(* IEC 61131-3 sources: FibonacciChallenge/Class/SafetyManager (part 3) *)

        pPDOElement^.PDO_ID                 := PDO_ID;
        pPDOElement^.Length                 := Length;
        pPDOElement^.ThisDomainsRole        := SourceDest_IsDest;

        pPDOElement^.SourceInfo.SafetyNbr   := 0;
        pPDOElement^.SourceInfo.DomainNr    := SourceDomain;
        pPDOElement^.SourceInfo.PathLen     := SourcePathLen;
        pPDOElement^.SourceInfo.pPath$pVoid := To_StdLib.Malloc(size:= SourcePathLen);
        if pPDOElement^.SourceInfo.pPath then
          _memcpy(ptr1:=pPDOElement^.SourceInfo.pPath, ptr2:=pSourcePath, cntr:=SourcePathLen);
        else
          LogError("@0464 (SafetyManager::IsAffectedByPDO) Failed to allocate memory for PDO path info");
          ClassState := -1;
          return;
        end_if;

        pPDOElement^.DestInfo.SafetyNbr     := pSafetyNbr^;
        pPDOElement^.DestInfo.DomainNr      := DestDomain;
        pPDOElement^.DestInfo.PathLen       := DestPathLen;
        pPDOElement^.DestInfo.pPath$pVoid   := To_StdLib.Malloc(size:= DestPathLen);
        if pPDOElement^.DestInfo.pPath then
          _memcpy(ptr1:=pPDOElement^.DestInfo.pPath, ptr2:=pDestPath, cntr:=DestPathLen);
        else
          LogError("@0464 (SafetyManager::IsAffectedByPDO) Failed to allocate memory for PDO path info");
          ClassState := -1;
          return;
        end_if;

        pPDOElement^.pSafety              := pDestSafety;

        // if we're the master, we may also route interfaceframes
        if IsInterfaceFrame then

          // search for the source of this PDO
          pHelpManaging := pFirstManagingInterfaceComponent;
          while pHelpManaging do
            if (To_StdLib.MemCmp(pHelpManaging^.pModulePath, pSourcePath, SourcePathLen) = 0) then
              exit;
            else
              pHelpManaging := pHelpManaging^.pNext;
            end_if;
          end_while;

          pPDOElement^.pManagingSource := pHelpManaging;
        end_if;

        if pPDOElement^.pManagingSource then

          // if the module is marked as optional and the PDO is not optional => the module is also not optional
          if pPDOElement^.pManagingSource^.InfoBits.IsOptional & (PDOInfo.IsOptional = FALSE) then
            pPDOElement^.pManagingSource^.InfoBits.IsOptional  := FALSE;
          end_if;

          // check if we can recycle the memory of another DO (if this data is already transferred to this managing module
          pRecyclePDO := CheckPDORecycle(SourceDest_IsSource, pPDOElement);

          // only if there is enough space or we already have a memory
          if pRecyclePDO | ((pPDOElement^.pManagingSource^.PDOReadMemUsed + pPDOElement^.Length) <= pPDOElement^.pManagingSource^.PDOReadMemAvailable) then
            if IsInterfaceFrame then
              pPDOElement^.SourceInfo.SafetyNbr   := (GetIFInfoByCRC(InterfaceCRC, #TempOffset, #TempLen))$HDINT;
              if TempLen = Length then
                // get the place in the memory of the source managing module
                pPDOElement^.SourceInfo.pPDOMem       := pPDOElement^.pManagingSource^.pPDOReadSpace + TempOffset;
                pPDOElement^.SourceInfo.pPDOMemDPRAM  := pPDOElement^.pManagingSource^.pPDOReadSpaceDPRAM + TempOffset;

                pPDOElement^.SourceInfo.HandlePDODPRAM := pPDOElement^.pManagingSource^.ud_HandlePDOReadSpaceDPRAM;
                pPDOElement^.SourceInfo.OffsetPDODPRAM := TempOffset;

                // if we need new memory, tell the managing module
                if (TempOffset + Length) > pPDOElement^.pManagingSource^.PDOReadMemUsed then
                  pPDOElement^.pManagingSource^.PDOReadMemUsed := TempOffset + Length;

                  MyPara.uiCmd := CMD_SM_PDO_MEM_USAGE_RD;
                  MyPara.aPara[0] := pPDOElement^.pManagingSource^.PDOReadMemUsed$DINT;
                  pPDOElement^.pManagingSource^.pThis^.NewInst(#MyPara, #MyResult);
                end_if;

                MyPara.uiCmd := CMD_SM_ADD_INPUT_PDO;
                MyPara.aPara[0] := pPDOElement^.SourceInfo.pPDOMem$DINT;
                MyPara.aPara[1] := pPDOElement^.SourceInfo.pPDOMemDPRAM$DINT;
                MyPara.aPara[2] := pPDOElement^.SourceInfo.SafetyNbr$DINT;
                MyPara.aPara[3] := Length;
                MyPara.aPara[4] := PDOInfo.IsOptional;
                MyPara.aPara[5] := pPDOElement^.SourceInfo.HandlePDODPRAM$DINT; // Needed for Payload Support
                MyPara.aPara[6] := pPDOElement^.SourceInfo.OffsetPDODPRAM$DINT; // Needed for Payload Support
                MyPara.aPara[7] := 0;// target offset (not necessary here)
                MyPara.aPara[8] := SM_IF_VALIDITY_MARK$DINT;
                MyPara.aPara[9] := TRUE;

                pDestSafety^.pThis^.NewInst(#MyPara, #MyResult);
              else
                LogError("@0469 (SafetyManager::IsAffectedByPDO) Length of interface frames doesn't match the local configuration");
              end_if;

            else
              if pRecyclePDO then
                pPDOElement^.SourceInfo.pPDOMem       := pRecyclePDO^.SourceInfo.pPDOMem;
                pPDOElement^.SourceInfo.pPDOMemDPRAM  := pRecyclePDO^.SourceInfo.pPDOMemDPRAM;
              else
                pPDOElement^.SourceInfo.pPDOMem       := pPDOElement^.pManagingSource^.pPDOReadSpace + pPDOElement^.pManagingSource^.PDOReadMemUsed;
                pPDOElement^.SourceInfo.pPDOMemDPRAM  := pPDOElement^.pManagingSource^.pPDOReadSpaceDPRAM + pPDOElement^.pManagingSource^.PDOReadMemUsed;

                // if we need new memory, tell the managing module
                pPDOElement^.pManagingSource^.PDOReadMemUsed += pPDOElement^.Length;

                MyPara.uiCmd := CMD_SM_PDO_MEM_USAGE_RD;
                MyPara.aPara[0] := pPDOElement^.pManagingSource^.PDOReadMemUsed$DINT;
                pPDOElement^.pManagingSource^.pThis^.NewInst(#MyPara, #MyResult);
              end_if;
            end_if;
          else
            // we add the memory anyway to show the user how much he would need
            pPDOElement^.pManagingSource^.PDOReadMemUsed += pPDOElement^.Length;

            MyPara.uiCmd := CMD_SM_PDO_MEM_USAGE_RD;
            MyPara.aPara[0] := pPDOElement^.pManagingSource^.PDOReadMemUsed$DINT;
            pPDOElement^.pManagingSource^.pThis^.NewInst(#MyPara, #MyResult);

            LogError("@046B (SafetyManager::IsAffectedByPDO) Not enough read memory to map all PDOs");
            return;
          end_if;
        else

          LogError("@046C (SafetyManager::IsAffectedByPDO) Couldn't find source managing module for PDO");
          return;
        end_if;

        PDOElementNo += 1;
      else
        pSourceDest^ := SourceDest_IsForwarder;

        // if source and destination are not in this domain, is it a bifurcation or a linear forwarding?
        pPDOElement^.PDO_ID                 := PDO_ID;
        pPDOElement^.Length                 := Length;
        pPDOElement^.ThisDomainsRole        := SourceDest_IsForwarder;

        pPDOElement^.SourceInfo.DomainNr    := SourceDomain;
        pPDOElement^.SourceInfo.PathLen     := SourcePathLen;
        pPDOElement^.SourceInfo.pPath$pVoid := To_StdLib.Malloc(size:= SourcePathLen);
        if pPDOElement^.SourceInfo.pPath then
          _memcpy(ptr1:=pPDOElement^.SourceInfo.pPath, ptr2:=pSourcePath, cntr:=SourcePathLen);
        else
          LogError("@0464 (SafetyManager::IsAffectedByPDO) Failed to allocate memory for PDO path info");
          ClassState := -1;
          return;
        end_if;

        pPDOElement^.DestInfo.DomainNr      := DestDomain;
        pPDOElement^.DestInfo.PathLen       := DestPathLen;
        pPDOElement^.DestInfo.pPath$pVoid   := To_StdLib.Malloc(size:= DestPathLen);
        if pPDOElement^.DestInfo.pPath then
          _memcpy(ptr1:=pPDOElement^.DestInfo.pPath, ptr2:=pDestPath, cntr:=DestPathLen);
        else
          LogError("@0464 (SafetyManager::IsAffectedByPDO) Failed to allocate memory for PDO path info");
          ClassState := -1;
          return;
        end_if;

        // initialize with invalid;
        CopyCmdIndex := -1;

        // if we're the master, we may also route interfaceframes
        if IsInterfaceFrame then

          // search for the source of this PDO
          pHelpManaging := pFirstManagingInterfaceComponent;
          while pHelpManaging do
            if (To_StdLib.MemCmp(pHelpManaging^.pModulePath, pSourcePath, SourcePathLen) = 0) then
              exit;
            else
              pHelpManaging := pHelpManaging^.pNext;
            end_if;
          end_while;

          pPDOElement^.pManagingSource := pHelpManaging;
        end_if;

        if pPDOElement^.pManagingSource then

          // if the module is marked as optional and the PDO is not optional => the module is also not optional
          if pPDOElement^.pManagingSource^.InfoBits.IsOptional & (PDOInfo.IsOptional = FALSE) then
            pPDOElement^.pManagingSource^.InfoBits.IsOptional  := FALSE;
          end_if;

          // check if we can recycle the memory of another DO (if this data is already transferred to this managing module
          pRecyclePDO := CheckPDORecycle(SourceDest_IsSource, pPDOElement);

          if pRecyclePDO | ((pPDOElement^.pManagingSource^.PDOReadMemUsed + pPDOElement^.Length) <= pPDOElement^.pManagingSource^.PDOReadMemAvailable) then
            if pRecyclePDO then
              pPDOElement^.SourceInfo.pPDOMem       := pRecyclePDO^.SourceInfo.pPDOMem;
              pPDOElement^.SourceInfo.pPDOMemDPRAM  := pRecyclePDO^.SourceInfo.pPDOMemDPRAM;
            else
              pPDOElement^.SourceInfo.pPDOMem       := pPDOElement^.pManagingSource^.pPDOReadSpace + pPDOElement^.pManagingSource^.PDOReadMemUsed;
              pPDOElement^.SourceInfo.pPDOMemDPRAM  := pPDOElement^.pManagingSource^.pPDOReadSpaceDPRAM + pPDOElement^.pManagingSource^.PDOReadMemUsed;
              pPDOElement^.pManagingSource^.PDOReadMemUsed += pPDOElement^.Length;

              MyPara.uiCmd := CMD_SM_PDO_MEM_USAGE_RD;
              MyPara.aPara[0] := pPDOElement^.pManagingSource^.PDOReadMemUsed$DINT;
              pPDOElement^.pManagingSource^.pThis^.NewInst(#MyPara, #MyResult);
            end_if;
          else
            // we add the memory anyway to show the user how much he would need
            pPDOElement^.pManagingSource^.PDOReadMemUsed += pPDOElement^.Length;

            MyPara.uiCmd := CMD_SM_PDO_MEM_USAGE_RD;
            MyPara.aPara[0] := pPDOElement^.pManagingSource^.PDOReadMemUsed$DINT;
            pPDOElement^.pManagingSource^.pThis^.NewInst(#MyPara, #MyResult);

            LogError("@046B (SafetyManager::IsAffectedByPDO) Not enough read memory to map all PDOs");
            return;
          end_if;
        else
          LogError("@046C (SafetyManager::IsAffectedByPDO) Couldn't find source managing module for PDO");
          return;
        end_if;

        // if we're the master, we may also route interfaceframes
        if IsInterfaceFrame then
          // search for the destination of this PDO
          pHelpManaging := pFirstManagingInterfaceComponent;
          while pHelpManaging do
            if (To_StdLib.MemCmp(pHelpManaging^.pModulePath, pDestPath, DestPathLen) = 0) then
              exit;
            else
              pHelpManaging := pHelpManaging^.pNext;
            end_if;
          end_while;

          pPDOElement^.pManagingDest := pHelpManaging;
        end_if;

        if pPDOElement^.pManagingDest then

          // if the module is marked as optional and the PDO is not optional => the module is also not optional
          if pPDOElement^.pManagingDest^.InfoBits.IsOptional & (PDOInfo.IsOptional = FALSE) then
            pPDOElement^.pManagingDest^.InfoBits.IsOptional  := FALSE;
          end_if;

          if pPDOElement^.pManagingDest = pPDOElement^.pManagingSource then
            LogError("@0470 (SafetyManager::IsAffectedByPDO) In PDO Forwarding a domain can't be the source and the destination!");
          end_if;

          // check if we can recycle the memory of another DO (if this data is already transferred to this managing module
          pRecyclePDO := CheckPDORecycle(SourceDest_IsDest, pPDOElement);

          if pRecyclePDO | ((pPDOElement^.pManagingDest^.PDOWriteMemUsed + pPDOElement^.Length) <= pPDOElement^.pManagingDest^.PDOWriteMemAvailable) then

            // if we can't use the copy command
            if b_SafetyOnLocalCDIAS then
              // remember the pointer to the memory to copy it manually in rt postscan method
              if pRecyclePDO then
                // this PDO is already in the memory of the managing node, we don't have to copy it again
                pPDOElement^.DestInfo.pPDOMem := NIL;//pRecyclePDO^.SourceInfo.pPDOMem;
              else
                pPDOElement^.DestInfo.pPDOMem := pPDOElement^.pManagingDest^.pPDOWriteSpace + pPDOElement^.pManagingDest^.PDOWriteMemUsed;
              end_if;
            else
              if pRecyclePDO then
                // this PDO is already in the memory of the managing node, we don't have to copy it again
                pPDOElement^.DestInfo.pPDOMemDPRAM := NIL;//pRecyclePDO^.DestInfo.pPDOMemDPRAM;
              else
                pPDOElement^.DestInfo.pPDOMemDPRAM := pPDOElement^.pManagingDest^.pPDOWriteSpaceDPRAM + pPDOElement^.pManagingDest^.PDOWriteMemUsed;
              end_if;

              CopyCmdIndex := GetNewMovDO();
              if CopyCmdIndex < 0 then
                pPDOElement^.DestInfo.pPDOMem := pPDOElement^.pManagingDest^.pPDOWriteSpace + pPDOElement^.pManagingDest^.PDOWriteMemUsed;
                LogError("@0465 (SafetyManager::IsAffectedByPDO) Failed to install copy command => PDO is beeing copied in RT");
              else
                aCopyCmds[CopyCmdIndex].pSettings^.ud_AddressDest := pPDOElement^.DestInfo.pPDOMemDPRAM$UDINT;
                aCopyCmds[CopyCmdIndex].pSettings^.ui_ByteCnt     := pPDOElement^.Length;
              end_if;
            end_if;

            // if we need new memory, tell the managing module
            if pRecyclePDO = NIL then
              pPDOElement^.pManagingDest^.PDOWriteMemUsed += pPDOElement^.Length;

              MyPara.uiCmd := CMD_SM_PDO_MEM_USAGE_WR;
              MyPara.aPara[0] := pPDOElement^.pManagingDest^.PDOWriteMemUsed$DINT;
              pPDOElement^.pManagingDest^.pThis^.NewInst(#MyPara, #MyResult);
            end_if;
          else
            // we add the memory anyway to show the user how much he would need
            pPDOElement^.pManagingDest^.PDOWriteMemUsed += pPDOElement^.Length;

            MyPara.uiCmd := CMD_SM_PDO_MEM_USAGE_WR;
            MyPara.aPara[0] := pPDOElement^.pManagingDest^.PDOWriteMemUsed$DINT;
            pPDOElement^.pManagingDest^.pThis^.NewInst(#MyPara, #MyResult);

            LogError("@0466 (SafetyManager::IsAffectedByPDO) Not enough write memory to map all PDOs");
            return;
          end_if;
        else
          LogError("@0467 (SafetyManager::IsAffectedByPDO) Couldn't find destination managing module for PDO");
          return;
        end_if;

        pPDOElement^.CopyCmdIndex := CopyCmdIndex;

        PDOElementNo += 1;
      end_if;

    end_if;
  end_if;

END_FUNCTION

FUNCTION SafetyManager::GetDestManagingOfDO
  VAR_INPUT
    pDO 	: ^SafetyCDIAS_Base::SDOHeader;
  END_VAR
  VAR_OUTPUT
    pDestManaging 	: ^t_ManagingComponent;
  END_VAR
  VAR
    pHelpManaging 	          : ^t_ManagingComponent;
    pAddDynSlaveRsp           : ^t_AddDynSlaveRsp;
    pRemDynSlaveRsp           : ^t_RemDynSlaveRsp;
    pHelpConfig               : ^t_CfgListElem;
    pHelpConnection           : ^t_FSoEConnectionDetails;
    MyPara                    : CmdStruct;
    MyResult                  : results;
    i                         : USINT;
    b_ConnectionAlreadyExists : BOOL;
  END_VAR

  pDestManaging := NIL;

  // maybe it's one of the interface domains
  pHelpManaging := pFirstManagingInterfaceComponent;
  while pHelpManaging do
    if (pHelpManaging^.FlexCon.SafetyNumber = pDO^.DstAdr) then
      if (pDO^.StdHeader.Typ.Response) & ((pDO^.StdHeader.Cmd = SM_SDO_COMMAND_ADD_DYN_SLAVE) | (pDO^.StdHeader.Cmd = SM_SDO_COMMAND_REMOVE_DYN_SLAVE)) then

        // if the initialisation of the class is not finished or failed
        if (sFlexCon.Role <> _NoFlexCon) & (ClassState <> 1) then
          // don't forward add or remove dyn slave requests. otherwise the order in the managing module is likely to be wrong if flexcon is used in combination with interface frames.
          return;
        end_if;

        if (pDO^.StdHeader.Cmd = SM_SDO_COMMAND_ADD_DYN_SLAVE) then
          pAddDynSlaveRsp := pDO$^t_AddDynSlaveRsp;

          // if it was successful and we have a safety host module pointer => try to install the PDO
          if (pAddDynSlaveRsp^.Retcode = 0) & sFlexCon.pSafetyHost then
#ifdef SAFETY_DEBUG_LOGGING_ACTIVATED
            LogError("@DBG AddDynSlave Response detected in SafetyManager of Host (succeeded)");
#endif

            // install the access to the next free memory on the VBC

            // we're the host => search for the FSoE connection with the host flags
            pHelpConfig := pConfigs;
            while pHelpConfig do
              pHelpConnection := pHelpConfig^.pFirstFSoEConnection;
              while pHelpConnection do
                if ((pHelpConnection^.Flags AND SM_FLAGS_FLEXCON_MASK) = SM_FLAGS_FLEXCON_HOST) &   // check if it's the right kind of connection
//                   (pHelpConnection^.InternalConnectionState =  FCS_RESET)               &          // check if it's still free
                   (pHelpConnection^.MasterReadOffset  = pAddDynSlaveRsp^.SafeOutOffset) &          // check if offsets and lengths match
                   (pHelpConnection^.MasterWriteOffset = pAddDynSlaveRsp^.SafeInOffset)  &
                   (pHelpConnection^.MasterReadSize    = pAddDynSlaveRsp^.SafeOutLength) &
                   (pHelpConnection^.MasterWriteSize   = pAddDynSlaveRsp^.SafeInLength) then

#ifdef SAFETY_DEBUG_LOGGING_ACTIVATED
                  LogValue(pString:="@DBG HOST: Found FSoE Connection of FlexConHost to install the cyclic PDO Routing between 0x{0} local and 0x{1} at Node", Value:=pHelpConnection^.OwnerSafetyNbr, Value2:=pHelpManaging^.FlexCon.SafetyNumber);
#endif

                  // remember if we already had this connection before
                  b_ConnectionAlreadyExists := pHelpManaging^.FlexCon.pCopyCmd <> NIL;

                  if b_ConnectionAlreadyExists = FALSE then
                    pHelpManaging^.FlexCon.WriteOffset:= pHelpManaging^.PDOWriteMemUsed$UINT;
                    pHelpManaging^.FlexCon.WriteLen   := pHelpConnection^.MasterReadSize;
                  end_if;

                  // GET THE DATA FROM THE SCP TO THE VBC

                  MyPara.uiCmd := CMD_SM_ADD_OUTPUT_PDO;
//                      MyPara.aPara[0] := 1;  not used // mark as interface frame PDO
                  sFlexCon.pSafetyHost^.pThis^.NewInst(#MyPara, #MyResult);

  //                  pPDOElement^.SourceInfo.pPDOMem       := MyResult.aData[0]$^USINT;
  //                  pPDOElement^.SourceInfo.pPDOMemDPRAM  := MyResult.aData[4]$^USINT;
  //                  pPDOElement^.SourceInfo.HandlePDODPRAM:= MyResult.aData[8]$UDINT;   // Needed for Payload Support
  //                  pPDOElement^.SourceInfo.OffsetPDODPRAM:= MyResult.aData[12]$UDINT;  // Needed for Payload Support

                  // check if we already have a copy pointer
                  if pHelpManaging^.FlexCon.pCopyCmd then
                    pHelpManaging^.FlexCon.pCopyCmd^.pSource  := MyResult.aData[0]$^USINT + pHelpConnection^.MasterReadOffset;
                    pHelpManaging^.FlexCon.pCopyCmd^.pDest    := pHelpManaging^.pPDOWriteSpace + pHelpManaging^.FlexCon.WriteOffset;
                    pHelpManaging^.FlexCon.pCopyCmd^.Size     := pHelpManaging^.FlexCon.WriteLen;
                  else
                    // create a new
                    if FSoECopyCmdNo < MAX_FSOE_CONNECTIONS then
                      aFSoECopyCmds[FSoECopyCmdNo].pSource  := MyResult.aData[0]$^USINT + pHelpConnection^.MasterReadOffset;
                      aFSoECopyCmds[FSoECopyCmdNo].pDest    := pHelpManaging^.pPDOWriteSpace + pHelpManaging^.FlexCon.WriteOffset;
                      aFSoECopyCmds[FSoECopyCmdNo].Size     := pHelpManaging^.FlexCon.WriteLen;
                      pHelpManaging^.FlexCon.pCopyCmd := #aFSoECopyCmds[FSoECopyCmdNo];
                      FSoECopyCmdNo                         += 1;
                    else
                      LogValue("@0493 (SafetyManager::GetDestManagingOfDO) Maximum limit of allowed FSoE connections exceeded (0x{0})", Value:=MAX_FSOE_CONNECTIONS);
                    end_if;
                  end_if;

                  if b_ConnectionAlreadyExists = FALSE then
                    pHelpManaging^.PDOWriteMemUsed += pHelpManaging^.FlexCon.WriteLen;
                    MyPara.uiCmd    := CMD_SM_PDO_MEM_USAGE_WR;
                    MyPara.aPara[0] := pHelpManaging^.PDOWriteMemUsed$DINT;
                    pHelpManaging^.pThis^.NewInst(#MyPara, #MyResult);

                    pHelpManaging^.FlexCon.ReadOffset := pHelpManaging^.PDOReadMemUsed$UINT;
                    pHelpManaging^.FlexCon.ReadLen    := pHelpConnection^.MasterWriteSize;
                  end_if;

                  // HOW TO GET DATA FROM THE VBC TO THE SCP

                  MyPara.uiCmd := CMD_SM_ADD_INPUT_PDO;
                  MyPara.aPara[0] := (pHelpManaging^.pPDOReadSpace + pHelpManaging^.FlexCon.ReadOffset)$DINT;
                  MyPara.aPara[1] := 0;
                  MyPara.aPara[2] := pHelpManaging^.FlexCon.SafetyNumber$DINT;
                  MyPara.aPara[3] := pHelpManaging^.FlexCon.ReadLen;
                  MyPara.aPara[4] := 0;
                  MyPara.aPara[5] := 0;
                  MyPara.aPara[6] := 0;
                  MyPara.aPara[7] := pHelpConnection^.MasterWriteOffset;
                  MyPara.aPara[8] := SM_IF_VALIDITY_MARK$DINT;
                  MyPara.aPara[9] := FALSE; // no interface frame => needed to reuse the same input PDO at the module

                  if sFlexCon.pSafetyHost^.pThis^.NewInst(#MyPara, #MyResult) = ERROR then
                    LogError(e_msg:="@05DE (SafetyManager::GetDestManagingOfDO) Failed to add FlexCon PDO to safe CPU PDO input buffer (Host side)");
                  end_if;

                  // check if we already have a input pdo pointer
                  if pHelpManaging^.FlexCon.pInputPdo then
                    pHelpManaging^.FlexCon.pInputPdo^.pSafety := sFlexCon.pSafetyHost;
                    pHelpManaging^.FlexCon.pInputPdo^.pMem    := MyPara.aPara[0];
                  else
                    if FSoEInputPDONo < MAX_FSOE_CONNECTIONS then
                      aFSoEInputPDOs[FSoEInputPDONo].pSafety    := sFlexCon.pSafetyHost;
                      aFSoEInputPDOs[FSoEInputPDONo].pMem       := MyPara.aPara[0];
                      pHelpManaging^.FlexCon.pInputPdo          := #aFSoEInputPDOs[FSoEInputPDONo];
                      FSoEInputPDONo += 1;
                    else
                      LogValue("@0490 (SafetyManager::GetDestManagingOfDO) Maximum limit of allowed FSoE input Frames exceeded (0x{0})", Value:=MAX_FSOE_CONNECTIONS);
                    end_if;
                  end_if;

#ifdef SAFETY_DEBUG_LOGGING_ACTIVATED
  #pragma message("RamAnd 20.11.2014 16:41 \ testweise mapping loggen")
                  LogValue("@DBG (SafetyManager::GetDestManagingOfDO) Mng => Modul: Wr Offset Modul: 0x{0}, Rd Offset Mng: 0x{1}, Größe: 0x{2}", Value:=pHelpConnection^.MasterWriteOffset, Value2:=pHelpManaging^.FlexCon.ReadOffset, Value3:=pHelpManaging^.FlexCon.ReadLen);
                  LogValue("@DBG (SafetyManager::GetDestManagingOfDO) Modul => Mng: Rd Offset Modul: 0x{0}, Wr Offset Mng: 0x{1}, Größe: 0x{2}", Value:=pHelpConnection^.MasterReadOffset, Value2:=pHelpManaging^.FlexCon.WriteOffset, Value3:=pHelpManaging^.FlexCon.WriteLen);
#endif

                  if b_ConnectionAlreadyExists = FALSE then
                    pHelpManaging^.PDOReadMemUsed += pHelpManaging^.FlexCon.ReadLen;

                    MyPara.uiCmd := CMD_SM_PDO_MEM_USAGE_RD;
                    MyPara.aPara[0] := pHelpManaging^.PDOReadMemUsed$DINT;
                    pHelpManaging^.pThis^.NewInst(#MyPara, #MyResult);
                  end_if;

                  // mark the connection as established
//                  pHelpConnection^.InternalConnectionState := FCS_CONNECTION;

                  // remember the connection if it's connected
                  pHelpManaging^.FlexCon.pFSoEConnection := pHelpConnection;

                  // we got our connection, stop cycling through the rest of the configurations
                  pDestManaging := pHelpManaging;
                  return;
                end_if;

                pHelpConnection := pHelpConnection^.pNext;
              end_while;
              pHelpConfig := pHelpConfig^.pNext;
            end_while;
          else
            LogValue(pString:="@05DF (SafetyManager::GetDestManagingOfDO) AddDynSlave Response detected in SafetyManager of Host (failed with retcode 0x{0})", Value:=pAddDynSlaveRsp^.Retcode);
          end_if;
        else
          pRemDynSlaveRsp := pDO$^t_RemDynSlaveRsp;

          if pRemDynSlaveRsp^.Retcode = 0 then
#ifdef SAFETY_DEBUG_LOGGING_ACTIVATED
            LogError("@DBG RemoveDynSlave Response detected in SafetyManager of Host (succeeded)");
#endif
            if pHelpManaging^.FlexCon.pFSoEConnection then
              // remove the InputPDO from the Safety CPU
              if pHelpManaging^.FlexCon.pInputPdo & pHelpManaging^.FlexCon.pInputPdo^.pMem & pHelpManaging^.FlexCon.pInputPdo^.pSafety then
                // unregister this PDO
                MyPara.uiCmd := CMD_SM_REMOVE_INPUT_PDO;
                MyPara.aPara[0] := pHelpManaging^.FlexCon.pInputPdo^.pMem;
                MyPara.aPara[1] := 0;
                pHelpManaging^.FlexCon.pInputPdo^.pSafety^.pThis^.NewInst(#MyPara, #MyResult);
              end_if;

//              pHelpManaging^.FlexCon.pFSoEConnection^.InternalConnectionState := FCS_RESET;
              pHelpManaging^.FlexCon.pFSoEConnection := NIL;
            end_if;
          else
            LogValue(pString:="@05E0 (SafetyManager::GetDestManagingOfDO) RemoveDynSlave Response detected in SafetyManager of Host (failed with retcode 0x{0})", Value:=pRemDynSlaveRsp^.Retcode);
          end_if;
        end_if;
      end_if;

      pDestManaging := pHelpManaging;
      return;
    end_if;

    if pHelpManaging^.ModuleNo then
      for i := 0 to (pHelpManaging^.ModuleNo-1) do
        if pHelpManaging^.ModuleInfo[i].SafetyNbr = pDO^.DstAdr then
          pDestManaging := pHelpManaging;
          return;
        end_if;
      end_for;
    end_if;

    pHelpManaging := pHelpManaging^.pNext;
  end_while;

END_FUNCTION

FUNCTION SafetyManager::GetDestSafetyOfDO
  VAR_INPUT
    pDO 	: ^SafetyCDIAS_Base::SDOHeader;
  END_VAR
  VAR_OUTPUT
    pDestSafety 	: ^t_SafetyComponent;
  END_VAR
  VAR
    pHelpSafety 	            : ^t_SafetyComponent;
    pAddDynSlaveRsp           : ^t_AddDynSlaveRsp;
    pRemDynSlaveRsp           : ^t_RemDynSlaveRsp;
    pHelpConfig               : ^t_CfgListElem;
    pHelpConnection           : ^t_FSoEConnectionDetails;
    MyPara                    : CmdStruct;
    MyResult                  : results;
    b_ConnectionAlreadyExists : BOOL;
  END_VAR

  pDestSafety := NIL;

  // check if it's a SDO addressed via safety number
  if (pDO^.StdHeader.Typ AND SSDO_MASK_TYPE) = FRM_TYPECODE_SSDO_MOD_TP then
    // we can't find it via Topology path
    LogError("@043C (SafetyManager::GetDestSafetyOfDO) Misdirected SDO via Topology path. Addressee can't be found here");
    return;
  end_if;

  pHelpSafety := pFirstSafetyComponent;
  while pHelpSafety do
    if pHelpSafety^.SafetyNbr = pDO^.DstAdr then

      // if it's a response to AddDynSlave or RemoveDynSlave request
      if (pDO^.StdHeader.Typ.Response) & ((pDO^.StdHeader.Cmd = SM_SDO_COMMAND_ADD_DYN_SLAVE) | (pDO^.StdHeader.Cmd = SM_SDO_COMMAND_REMOVE_DYN_SLAVE)) then

        // if the initialisation of the class is not finished or failed
        if (sFlexCon.Role <> _NoFlexCon) & (ClassState <> 1) then
          // don't forward add or remove dyn slave requests. otherwise the order in the managing module is likely to be wrong if flexcon is used in combination with interface frames.
          return;
        end_if;

        // if it's an AddDynSlave response
        if (pDO^.StdHeader.Cmd = SM_SDO_COMMAND_ADD_DYN_SLAVE) then
          pAddDynSlaveRsp := pDO$^t_AddDynSlaveRsp;

          // if it was successful and we have a safety host managing module pointer as well as a safety number connected with it => try to install the PDO
          if (pAddDynSlaveRsp^.Retcode = 0) & sFlexCon.pManaging2Host & sFlexCon.pManaging2Host^.FlexCon.SafetyNumber then
#ifdef SAFETY_DEBUG_LOGGING_ACTIVATED
            LogError("@DBG AddDynSlave Response detected in SafetyManager of Node (succeeded)");
#endif

            // install the access to the next free memory on the VBC

            // we're the node => search for the FSoE connection with the node flags
            pHelpConfig := pConfigs;
            while pHelpConfig do
              pHelpConnection := pHelpConfig^.pFirstFSoEConnection;
              while pHelpConnection do
                if ((pHelpConnection^.Flags AND SM_FLAGS_FLEXCON_MASK) = SM_FLAGS_FLEXCON_NODE) & // check if it's the right kind of connection
                    (pHelpConnection^.MasterWriteSize   = pAddDynSlaveRsp^.SafeOutLength) &
                    (pHelpConnection^.MasterReadSize    = pAddDynSlaveRsp^.SafeInLength) then

#ifdef SAFETY_DEBUG_LOGGING_ACTIVATED
                  LogValue(pString:="@DBG NODE: Found FSoE Connection of FlexConNode to install the cyclic PDO Routing between 0x{0} local and 0x{1} at Host", Value:=pHelpConnection^.OwnerSafetyNbr, Value2:=sFlexCon.pManaging2Host^.FlexCon.SafetyNumber);
#endif

                  // remember if we already had this connection before
                  b_ConnectionAlreadyExists := sFlexCon.pManaging2Host^.FlexCon.pCopyCmd <> NIL;

                  // if we just created this connection
                  if b_ConnectionAlreadyExists = FALSE then
                    // remember offset and length of the write access
                    sFlexCon.pManaging2Host^.FlexCon.WriteOffset:= sFlexCon.pManaging2Host^.PDOWriteMemUsed$UINT;
                    sFlexCon.pManaging2Host^.FlexCon.WriteLen   := pAddDynSlaveRsp^.SafeOutLength;
                  end_if;

                  // GET THE DATA FROM THE SCP TO THE VBC

                  MyPara.uiCmd := CMD_SM_ADD_OUTPUT_PDO;
//                      MyPara.aPara[0] := 1;  not used // mark as interface frame PDO
                  pHelpSafety^.pThis^.NewInst(#MyPara, #MyResult);

  //                  pPDOElement^.SourceInfo.pPDOMem       := MyResult.aData[0]$^USINT;
  //                  pPDOElement^.SourceInfo.pPDOMemDPRAM  := MyResult.aData[4]$^USINT;
  //                  pPDOElement^.SourceInfo.HandlePDODPRAM:= MyResult.aData[8]$UDINT;   // Needed for Payload Support
  //                  pPDOElement^.SourceInfo.OffsetPDODPRAM:= MyResult.aData[12]$UDINT;  // Needed for Payload Support

                  // check if we already have a copy pointer
                  if sFlexCon.pManaging2Host^.FlexCon.pCopyCmd then
                    sFlexCon.pManaging2Host^.FlexCon.pCopyCmd^.pSource  := MyResult.aData[0]$^USINT + pHelpConnection^.SlaveReadOffset;
                    sFlexCon.pManaging2Host^.FlexCon.pCopyCmd^.pDest    := sFlexCon.pManaging2Host^.pPDOWriteSpace + sFlexCon.pManaging2Host^.FlexCon.WriteOffset;
                    sFlexCon.pManaging2Host^.FlexCon.pCopyCmd^.Size     := sFlexCon.pManaging2Host^.FlexCon.WriteLen;
                  else
                    if FSoECopyCmdNo < MAX_FSOE_CONNECTIONS then
                      aFSoECopyCmds[FSoECopyCmdNo].pSource  := MyResult.aData[0]$^USINT + pHelpConnection^.SlaveReadOffset;
                      aFSoECopyCmds[FSoECopyCmdNo].pDest    := sFlexCon.pManaging2Host^.pPDOWriteSpace + sFlexCon.pManaging2Host^.FlexCon.WriteOffset;
                      aFSoECopyCmds[FSoECopyCmdNo].Size     := sFlexCon.pManaging2Host^.FlexCon.WriteLen;
                      sFlexCon.pManaging2Host^.FlexCon.pCopyCmd := #aFSoECopyCmds[FSoECopyCmdNo];
                      FSoECopyCmdNo                         += 1;
                    else
                      LogValue("@0493 (SafetyManager::GetDestSafetyOfDO) Maximum limit of allowed FSoE connections exceeded (0x{0})", Value:=MAX_FSOE_CONNECTIONS);
                    end_if;
                  end_if;

                  // if we just created this connection
                  if b_ConnectionAlreadyExists = FALSE then
                    // increase the used write memory on the managing module
                    sFlexCon.pManaging2Host^.PDOWriteMemUsed += sFlexCon.pManaging2Host^.FlexCon.WriteLen;

                    MyPara.uiCmd    := CMD_SM_PDO_MEM_USAGE_WR;
                    MyPara.aPara[0] := sFlexCon.pManaging2Host^.PDOWriteMemUsed$DINT;
                    sFlexCon.pManaging2Host^.pThis^.NewInst(#MyPara, #MyResult);

                    // remember offset and length of the read access
                    sFlexCon.pManaging2Host^.FlexCon.ReadOffset:= sFlexCon.pManaging2Host^.PDOReadMemUsed$UINT;
                    sFlexCon.pManaging2Host^.FlexCon.ReadLen   := pHelpConnection^.MasterReadSize;
                  end_if;

                  // HOW TO GET DATA FROM THE VBC TO THE SCP

                  MyPara.uiCmd := CMD_SM_ADD_INPUT_PDO;
                  MyPara.aPara[0] := (sFlexCon.pManaging2Host^.pPDOReadSpace + sFlexCon.pManaging2Host^.FlexCon.ReadOffset)$DINT;
                  MyPara.aPara[1] := 0;
                  MyPara.aPara[2] := sFlexCon.pManaging2Host^.FlexCon.SafetyNumber$DINT;
                  MyPara.aPara[3] := sFlexCon.pManaging2Host^.FlexCon.ReadLen;
                  MyPara.aPara[4] := 0;
                  MyPara.aPara[5] := 0;
                  MyPara.aPara[6] := 0;
                  MyPara.aPara[7] := pHelpConnection^.SlaveWriteOffset;
                  MyPara.aPara[8] := SM_IF_VALIDITY_MARK$DINT;
                  MyPara.aPara[9] := FALSE; // no interface frame => needed to reuse the same input PDO at the module

                  if pHelpSafety^.pThis^.NewInst(#MyPara, #MyResult) = ERROR then
                    LogError(e_msg:="@05E1 (SafetyManager::GetDestManagingOfDO) Failed to add FlexCon PDO to safe CPU PDO input buffer (Node side)");
                  end_if;

                  // check if we already have a input pdo pointer
                  if sFlexCon.pManaging2Host^.FlexCon.pInputPdo then
                    sFlexCon.pManaging2Host^.FlexCon.pInputPdo^.pSafety := pHelpSafety;
                    sFlexCon.pManaging2Host^.FlexCon.pInputPdo^.pMem    := MyPara.aPara[0];
                  else
                    if FSoEInputPDONo < MAX_FSOE_CONNECTIONS then
                      aFSoEInputPDOs[FSoEInputPDONo].pSafety    := pHelpSafety;
                      aFSoEInputPDOs[FSoEInputPDONo].pMem       := MyPara.aPara[0];
                      sFlexCon.pManaging2Host^.FlexCon.pInputPdo := #aFSoEInputPDOs[FSoEInputPDONo];
                      FSoEInputPDONo += 1;
                    else
                      LogValue("@0490 (SafetyManager::GetDestSafetyOfDO) Maximum limit of allowed FSoE input Frames exceeded (0x{0})", Value:=MAX_FSOE_CONNECTIONS);
                    end_if;
                  end_if;

#ifdef SAFETY_DEBUG_LOGGING_ACTIVATED
  #pragma message("RamAnd 20.11.2014 16:41 \ testweise mapping loggen")
                  LogValue("@DBG (SafetyManager::GetDestSafetyOfDO) Mng => Modul: Wr Offset Modul: 0x{0}, Rd Offset Mng: 0x{1}, Größe: 0x{2}", Value:=pHelpConnection^.SlaveWriteOffset, Value2:=sFlexCon.pManaging2Host^.FlexCon.ReadOffset, Value3:=sFlexCon.pManaging2Host^.FlexCon.ReadLen);
                  LogValue("@DBG (SafetyManager::GetDestSafetyOfDO) Modul => Mng: Rd Offset Modul: 0x{0}, Wr Offset Mng: 0x{1}, Größe: 0x{2}", Value:=pHelpConnection^.SlaveReadOffset, Value2:=sFlexCon.pManaging2Host^.FlexCon.WriteOffset, Value3:=sFlexCon.pManaging2Host^.FlexCon.WriteLen);
#endif

                  // if we just created this connection
                  if b_ConnectionAlreadyExists = FALSE then
                    // increase the used read memory on the managing module
                    sFlexCon.pManaging2Host^.PDOReadMemUsed += sFlexCon.pManaging2Host^.FlexCon.ReadLen;

                    MyPara.uiCmd := CMD_SM_PDO_MEM_USAGE_RD;
                    MyPara.aPara[0] := sFlexCon.pManaging2Host^.PDOReadMemUsed$DINT;
                    sFlexCon.pManaging2Host^.pThis^.NewInst(#MyPara, #MyResult);
                  end_if;

                  // remember the connection if it's connected
                  sFlexCon.pManaging2Host^.FlexCon.pFSoEConnection := pHelpConnection;

                  // we got our connection, stop cycling through the rest of the configurations
                  pDestSafety := pHelpSafety;
                  return;
                end_if;

                pHelpConnection := pHelpConnection^.pNext;
              end_while;
              pHelpConfig := pHelpConfig^.pNext;
            end_while;
          else
            LogValue(pString:="@05E2 (SafetyManager::GetDestSafetyOfDO) AddDynSlave Response detected in SafetyManager of Node (failed with retcode 0x{0})", Value:=pAddDynSlaveRsp^.Retcode);
          end_if;
        else
          // it's a RemoveDynSlave response

          pRemDynSlaveRsp := pDO$^t_RemDynSlaveRsp;

          if pRemDynSlaveRsp^.Retcode = 0 then
#ifdef SAFETY_DEBUG_LOGGING_ACTIVATED
            LogError("@DBG RemoveDynSlave Response detected in SafetyManager of Node (succeeded)");
#endif

            if sFlexCon.pManaging2Host & sFlexCon.pManaging2Host^.FlexCon.pFSoEConnection then
              // remove the InputPDO from the Safety CPU
              if sFlexCon.pManaging2Host^.FlexCon.pInputPdo & sFlexCon.pManaging2Host^.FlexCon.pInputPdo^.pMem & sFlexCon.pManaging2Host^.FlexCon.pInputPdo^.pSafety then
                // unregister this PDO
                MyPara.uiCmd := CMD_SM_REMOVE_INPUT_PDO;
                MyPara.aPara[0] := sFlexCon.pManaging2Host^.FlexCon.pInputPdo^.pMem;
                MyPara.aPara[1] := 0;
                sFlexCon.pManaging2Host^.FlexCon.pInputPdo^.pSafety^.pThis^.NewInst(#MyPara, #MyResult);
              end_if;

//              sFlexCon.pManaging2Host^.FlexCon.pFSoEConnection^.InternalConnectionState := FCS_RESET;
              sFlexCon.pManaging2Host^.FlexCon.pFSoEConnection := NIL;
            end_if;

          else
            LogValue(pString:="@05E3 (SafetyManager::GetDestSafetyOfDO) RemoveDynSlave Response detected in SafetyManager of Node (failed with retcode 0x{0})", Value:=pRemDynSlaveRsp^.Retcode);
          end_if;
        end_if;
      end_if;

      pDestSafety := pHelpSafety;
      return;
    end_if;

    pHelpSafety := pHelpSafety^.pNext;
  end_while;

END_FUNCTION

FUNCTION VIRTUAL GLOBAL SafetyManager::RtWork
  VAR_INPUT
    EAX 	: UDINT;
  END_VAR
  VAR_OUTPUT
    state (EAX) 	: UDINT;
  END_VAR
  VAR
    i                 : UDINT;
    pPDOElement       : ^t_PDOElement;
    pFSoEElement      : ^t_FSoECopyCmd;
    AllCopyCmdsReady  : BOOL;
  END_VAR

  if EAX = CALL_OPTION_RT_PRESCAN then
    // prescan

//=================================================================================================
#ifdef VM_CLASS_TIME_MEASUREMENT
  StartTimeMeasurement(VARANTIME_RT);
#endif
//=================================================================================================

    // copy commands for udp connections (receiving via udp)
    if sUdpVars.ReceiveCopyCmdNo then
      // we may have some udp send data, so we better protect the copy mechanism
      UdpReceiveData.SectionStart();

      pFSoEElement := #sUdpVars.aReceiveCopyCmds[0];
      for i := 1 to sUdpVars.ReceiveCopyCmdNo do
        _memcpy(ptr1:=pFSoEElement^.pDest, ptr2:=pFSoEElement^.pSource, cntr:=pFSoEElement^.Size);
        pFSoEElement += sizeof(t_FSoECopyCmd);
      end_for;

      UdpReceiveData.SectionStop();
    end_if;

    case InitSSW of
//**********************************************************************************************************************************************************
      _Wait4CopyCmdStart:
        // start all used copy commands
        AllCopyCmdsReady := TRUE;
        if CopyCmdsUsed then
          for i := 0 to (CopyCmdsUsed-1) do
            if aCopyCmds[i].b_Ready4Action then
              aCopyCmds[i].pHandle^.ucCtrlStat := VARAN_DO_CONT_RUN;
            else
              AllCopyCmdsReady := FALSE;
              bd_LogRtMessagesInCy.UnkownCopySource := TRUE;
            end_if;
          end_for;
        end_if;

        if AllCopyCmdsReady then
          InitSSW := _FinishInitialisation;
        end_if;

//**********************************************************************************************************************************************************
      _InitFinished:
        // if we're master or we're actually time synchronizing
        if b_NewSyncMode & b_CheckTimeSyncTimeout then
          if (ops.tAbsolute - TimeSyncTimeStamp) > TIMESYNC_TIMEOUT then
            // increment timeout counter => message is shown in cyclic after x consecutive
            SyncTimeoutCounter += 1;
            b_CheckTimeSyncTimeout := FALSE; // => show Trace Message only once per error
            // restart the synchronisation (maybe the other domain has been disconnected)
            b_StartTimeSync := TRUE;
          end_if;
        end_if;

//**********************************************************************************************************************************************************
    end_case;

    // marker is set in cyclic priority (except on timeout), but time synchronisation has to be done in rt priority => start it from here
    if b_StartTimeSync then
      b_StartTimeSync := FALSE;

      StartTimeSync();
    end_if;

//=================================================================================================
#ifdef VM_CLASS_TIME_MEASUREMENT
  StopTimeMeasurement(VARANTIME_RT);
#endif
//=================================================================================================

  else
    // postscan

//=================================================================================================
#ifdef VM_CLASS_TIME_MEASUREMENT
  StartTimeMeasurement(VARANTIME_RTPOSTSCAN);
#endif
//=================================================================================================

    // copy data from our memory to the memory of the next domain
    if PDOElementNo then
      pPDOElement := #aPDOElements[0];
      for i := 1 to PDOElementNo do
        if (pPDOElement^.ThisDomainsRole = SourceDest_IsSource) |
           (pPDOElement^.ThisDomainsRole = SourceDest_IsForwarder) then
          if pPDOElement^.DestInfo.pPDOMem & pPDOElement^.SourceInfo.pPDOMem & pPDOElement^.Length then
            _memcpy(ptr1:=pPDOElement^.DestInfo.pPDOMem, ptr2:=pPDOElement^.SourceInfo.pPDOMem, cntr:=pPDOElement^.Length);
          end_if;
        end_if;
        pPDOElement += sizeof(t_PDOElement);
      end_for;
    elsif FSoECopyCmdNo then
      pFSoEElement := #aFSoECopyCmds[0];
      for i := 1 to FSoECopyCmdNo do
        _memcpy(ptr1:=pFSoEElement^.pDest, ptr2:=pFSoEElement^.pSource, cntr:=pFSoEElement^.Size);
        pFSoEElement += sizeof(t_FSoECopyCmd);
      end_for;
    end_if;

    // copy commands for udp connections (sending via udp)
    if sUdpVars.SendCopyCmdNo then
      // we may have some udp send data, so we better protect the copy mechanism
      UdpSendData.SectionStart();

      pFSoEElement := #sUdpVars.aSendCopyCmds[0];
      for i := 1 to sUdpVars.SendCopyCmdNo do
        _memcpy(ptr1:=pFSoEElement^.pDest, ptr2:=pFSoEElement^.pSource, cntr:=pFSoEElement^.Size);
        pFSoEElement += sizeof(t_FSoECopyCmd);
      end_for;

      UdpSendData.SectionStop();
    end_if;

//=================================================================================================
#ifdef VM_CLASS_TIME_MEASUREMENT
  StopTimeMeasurement(VARANTIME_RTPOSTSCAN);
#endif
//=================================================================================================

  end_if;

#ifdef SAFETY_DEBUG_LOGGING_ACTIVATED
  if InitSSW <> OldInitSSW then
#ifdef SAFETY_DEBUG_TRACING_ACTIVATED
    LogValue("@DBG (SafetyManager::RtWork) InitSSW changed from {0} to {1}", Value:=OldInitSSW, Value2:=InitSSW);
#endif
    LogBuf[ActLogIndex].NewState := InitSSW;
    LogBuf[ActLogIndex].OldState := OldInitSSW;
    LogBuf[ActLogIndex].Command := 0;
    LogBuf[ActLogIndex].TimeSinceLastLog_us := OS_READMICROSEC();
    LogBuf[ActLogIndex].TimeSinceLastLog_us -= TimeStampLastLog_us;
    TimeStampLastLog_us := OS_READMICROSEC();
    if ActLogIndex = (LogBufferSize - 1) then
      ActLogIndex := 0;
    else
      ActLogIndex += 1;
    end_if;
  end_if;
  OldInitSSW := InitSSW;
#endif

  state := READY;

END_FUNCTION

FUNCTION SafetyManager::CheckTopSDO
  VAR_INPUT
    pPara 	: ^CmdStruct;
  END_VAR
  VAR
    pDO 	            : ^SafetyCDIAS_Base::SDOHeader;
    pCompDestPath     : ^USINT;
    pHelpConfig       : ^t_CfgListElem;
    pHelpSlave        : ^t_SlaveListElem;
    pHelpModule       : ^t_ModuleListElem;
    pHelpPdo          : ^t_PdoListElem;
    pHelpManaging     : ^t_ManagingComponent;
    pHelpSafety       : ^t_SafetyComponent;
    pHelpConnection   : ^t_FSoEConnectionDetails;
    MyPara            : CmdStruct;
    MyResult          : results;
    pTempMem          : ^USINT;
    pHelp             : ^USINT;
    TmpLen            : UINT;
    DomainChangeFound : BOOL;
    i                 : UDINT;
    DestDomain        : USINT;
    InterfaceCRC      : HDINT;
    TargetSafetyNbr   : HDINT;
    pActConnection    : ^t_UdpConnection;
    IPAddr            : HDINT;
  END_VAR

  // get a pointer to the compressed destination path
  pDO := (pPara^.aPara[1])$^SafetyCDIAS_Base::SDOHeader;
  pCompDestPath := (#pDO^.DstAdr)$^USINT;

  // if we have interfaceframes, check them first
  if pFirstManagingInterfaceComponent & (pCompDestPath^ = INTERFACE_CRC_MODE) then
    // after the mode byte we find the interface CRC
    InterfaceCRC := ((pCompDestPath + 1)$^HDINT)^;

    // if we have local connections and the source is not local => check the local connections for a receiver
    if pSortedConnections & (pPara^.aPara[2] <> this$DINT) then
      // we have to search for a receiver
      pHelpConnection := pSortedConnections;

      while pHelpConnection do
        if pHelpConnection^.SlavePathCompLen & pHelpConnection^.pSlavePathComp then
          if (pHelpConnection^.pSlavePathComp$^HDINT + 1)^ = InterfaceCRC then
            // we found the interface CRC, now we have to make a connection via the SafetyNumber between the actual config and the module handles
            pHelpSafety := pFirstSafetyComponent;
            while pHelpSafety do
              // we compare the safety number
              if pHelpSafety^.SafetyNbr = pHelpConnection^.OwnerSafetyNbr then
                // change the command, because now we forward it to the receiver
                pPara^.uiCmd := CMD_SM_SDO_TO_MODULE;

                pHelpSafety^.pThis^.NewInst(pPara, #MyResult);

                return;
              end_if;

              pHelpSafety := pHelpSafety^.pNext;
            end_while;
          end_if;
        end_if;

        pHelpConnection := pHelpConnection^.pNext;
      end_while;
    end_if;

    // if there are FSoE Connection
    if IFFSoENo then
      // if this system is the sender
      if (pPara^.aPara[2] = this$DINT) then
        // check the FSoE Connections
        for i := 0 to (IFFSoENo-1) do
          if aIFFSoEInfos[i].FromOtherSide.InterfaceCRC = InterfaceCRC then
            if aIFFSoEInfos[i].pManaging & aIFFSoEInfos[i].pManaging^.InfoBits.IsSynchron then
              aIFFSoEInfos[i].pManaging^.pThis^.NewInst(pPara, #MyResult);
            end_if;

            // we're done here
            return;
          end_if;
        end_for;

        // check if it's a local interface frame
        pHelpSafety := NIL;
        if LocalIFNo then
          for i := 0 to (LocalIFNo-1) do
            if aLocalIFs[i].InterfaceCRC = InterfaceCRC then
              // found it
              pHelpSafety := aLocalIFs[i].pSafetyModule;
              exit;
            end_if;
          end_for;
        end_if;

        if pHelpSafety then
          // change the command, because now we forward it to the receiver
          pPara^.uiCmd := CMD_SM_SDO_TO_MODULE;

          pHelpSafety^.pThis^.NewInst(pPara, #MyResult);
        else
          LogError("@043E (SafetyManager::CheckTopSDO) Couldn't find target of SDO via TOP (Interface Frame in FSoE mode)");
          LogValue("SrcAddr: {0} / InterfaceCRC: {1}", Value:=pDO^.SrcAdr, Value2:=InterfaceCRC);
        end_if;
      else
        // we have to search for a receiver
        pHelpConfig := pConfigs;
        while pHelpConfig do
          pHelpConnection := pHelpConfig^.pFirstFSoEConnection;
          while pHelpConnection do
            if pHelpConnection^.SlavePathCompLen & pHelpConnection^.pSlavePathComp then
              if (pHelpConnection^.pSlavePathComp$^HDINT + 1)^ = InterfaceCRC then
                // we found the interface CRC, now we have to make a connection via the SafetyNumber between the actual config and the module handles
                pHelpSafety := pFirstSafetyComponent;
                while pHelpSafety do
                  // we compare the safety number
                  if pHelpSafety^.SafetyNbr = pHelpConfig^.SafetyNbr then
                    // change the command, because now we forward it to the receiver
                    pPara^.uiCmd := CMD_SM_SDO_TO_MODULE;

                    pHelpSafety^.pThis^.NewInst(pPara, #MyResult);

                    return;
                  end_if;

                  pHelpSafety := pHelpSafety^.pNext;
                end_while;
              end_if;
            end_if;

            pHelpConnection := pHelpConnection^.pNext;
          end_while;
          pHelpConfig := pHelpConfig^.pNext;
        end_while;
      end_if;
    else
      if b_GotFSoEModules then
        // search in the module lists
        pHelpConfig := pConfigs;
        TargetSafetyNbr := 0;
        while pHelpConfig do
          pHelpModule := pHelpConfig^.pFirstModuleCfg;
          while pHelpModule do
            if pHelpModule^.ModuleInfo.InterfaceCRC = InterfaceCRC then
              TargetSafetyNbr := pHelpModule^.ModuleInfo.SafetyNbr;
            end_if;

            // if we found our target => forward the SDO to it
            if TargetSafetyNbr then
              pHelpSafety := pFirstSafetyComponent;
              while pHelpSafety do
                // we compare the safety number
                if pHelpSafety^.SafetyNbr = TargetSafetyNbr then
                  // change the command, because now we forward it to the receiver
                  pPara^.uiCmd := CMD_SM_SDO_TO_MODULE;

                  pHelpSafety^.pThis^.NewInst(pPara, #MyResult);

                  return;
                end_if;

                pHelpSafety := pHelpSafety^.pNext;
              end_while;
            end_if;

            pHelpModule := pHelpModule^.pNext;
          end_while;

          pHelpConfig := pHelpConfig^.pNext;
        end_while;
      else
  // check if we have an interface frame with this CRC
        pHelpConfig := pConfigs;
        while pHelpConfig do
          pHelpPdo := pHelpConfig^.pFirstPdoCfg;
          while pHelpPdo do
            // don't look at IFBroatCast PDOs, they are not distributed
            if (pHelpPdo^.PdoInfo.InterfaceCRC = InterfaceCRC) then
              if (pHelpPdo^.PdoInfo.Info.IFBroadCast = FALSE) then

                // if we found the CRC, forward it to the source of the PDO (the destination asks for the safety number)

                // check the source

                // if the master itself is the caller, it's from this system (check if it's for another system)
                if (pPara^.aPara[2] = this$DINT) then
                  pHelpManaging := pFirstManagingInterfaceComponent;
                  while pHelpManaging do
                    if (To_StdLib.MemCmp(pHelpManaging^.pModulePath, pHelpPdo^.PdoInfo.pSourcePath, pHelpPdo^.PdoInfo.SourcePathLen) = 0) then
                      exit;
                    else
                      pHelpManaging := pHelpManaging^.pNext;
                    end_if;
                  end_while;

                  if pHelpManaging then
                    if pHelpManaging^.InfoBits.IsSynchron then
                      pHelpManaging^.pThis^.NewInst(pPara, #MyResult);
                    end_if;
                  else
                    // no managing module found => continue search in our special safety module list
                    pHelpSafety := NIL;
                    if LocalIFNo then
                      for i := 0 to (LocalIFNo-1) do
                        if aLocalIFs[i].InterfaceCRC = InterfaceCRC then
                          // found it
                          pHelpSafety := aLocalIFs[i].pSafetyModule;
                          exit;
                        end_if;
                      end_for;
                    end_if;

                    if pHelpSafety then
                      // change the command, because now we forward it to the receiver
                      pPara^.uiCmd := CMD_SM_SDO_TO_MODULE;

                      pHelpSafety^.pThis^.NewInst(pPara, #MyResult);
                    else
                      // check the slave modules if there is one with the interface frame we need
                      pHelpConfig := pConfigs;
                      while pHelpConfig do
                        pHelpSlave := pHelpConfig^.pFirstSlaveCfg;
                        while pHelpSlave do

                          if (pHelpSlave^.SlaveInfo.Info.IsInterface) & (pHelpSlave^.SlaveInfo.InterfaceCRC = InterfaceCRC) then
                            // we have to add some additional information to the message

                            (*
                              Memory structure:
                                1 Byte destination domain
                                1 Byte IsInterfaceFrame (0/1)
                                2 Byte length of uncompressed path
                                x Byte uncompressed path
                                x Byte SDO message
                            *)

                            MyPara.uiCmd := CMD_SM_TOP_SDO_TO_MODULE;
                            MyPara.aPara[0] := sizeof(USINT) + sizeof(BOOL) + sizeof(UINT) + pHelpSlave^.SlaveInfo.PathLen + pPara^.aPara[0];

                            if ud_SizeTempMemCy >= MyPara.aPara[0]$UDINT then
                              pTempMem := pTempMemCy$^USINT;
                            else
                              LogError("@0440 (SafetyManager::CheckTopSDO) Temporary memory for cyclic task is too small!");
                              LogValue("AvaliableMem: {0} / NeededMem: {1}", Value:=ud_SizeTempMemCy, Value2:=MyPara.aPara[0]$UDINT);
                              return;
                            end_if;

                            TmpLen := pHelpSlave^.SlaveInfo.PathLen; // save some time with this local variable
                            DomainChangeFound := FALSE;
                            pHelp := pHelpSlave^.SlaveInfo.pPath + TmpLen - 2; // pointer on penultimate byte of path
                            // search from the end for the last domain change
                            for i := (TmpLen-2) to 3 by -1 do
                              if pHelp^ = HWT_ESCAPE_DOMAIN then
                                DomainChangeFound := TRUE;
                                DestDomain := (pHelp + 1)^;
                                exit;
                              end_if;

                              pHelp -= sizeof(USINT);
                            end_for;

                            // if there was no domainchange
                            if DomainChangeFound = FALSE then
                              // the master is the Dest
                              DestDomain := (pHelpSlave^.SlaveInfo.pPath + 2)^;
                            end_if;

                            pHelp := pTempMem;

                            // destination domain
                            pHelp^ := DestDomain;
                            pHelp += sizeof(USINT);

                            // is it for an interface frame?
                            pHelp^$BOOL := TRUE;
                            pHelp += sizeof(BOOL);

                            // length of uncompressed path
                            pHelp^$UINT := TmpLen;
                            pHelp += sizeof(UINT);

                            // uncompressed path
                            _memcpy(ptr1:=pHelp, ptr2:=pHelpSlave^.SlaveInfo.pPath, cntr:=TmpLen);
                            pHelp += TmpLen;

                            // SDO message
                            _memcpy(ptr1:=pHelp, ptr2:=pDO, cntr:=pPara^.aPara[0]$UDINT);

                            MyPara.aPara[1] := pTempMem$DINT;

                            NewInst(#MyPara, #MyResult);

                            // path can exist only once in a system
                            return;
                          end_if;

                          pHelpSlave := pHelpSlave^.pNext;
                        end_while;

                        pHelpConfig := pHelpConfig^.pNext;
                      end_while;

                      LogError("@0441 (SafetyManager::CheckTopSDO) Couldn't find target of SDO via TOP (Interface Frame)");
                      LogValue("SrcAddr: {0} / InterfaceCRC: {1}", Value:=pDO^.SrcAdr, Value2:=InterfaceCRC);
                    end_if;
                  end_if;
                else
                  // we got it from another system => check our modules
                  pHelpSafety := NIL;
                  if LocalIFNo then
                    for i := 0 to (LocalIFNo-1) do
                      if aLocalIFs[i].InterfaceCRC = InterfaceCRC then
                        // found it
                        pHelpSafety := aLocalIFs[i].pSafetyModule;
                        exit;
                      end_if;
                    end_for;
                  end_if;

                  if pHelpSafety then
                    // change the command, because now we forward it to the receiver
                    pPara^.uiCmd := CMD_SM_SDO_TO_MODULE;

                    pHelpSafety^.pThis^.NewInst(pPara, #MyResult);
                  else
                    LogError("@0441 (SafetyManager::CheckTopSDO) Couldn't find target of SDO via TOP (Interface Frame) received by another PLC");
                    LogValue("SrcAddr: {0} / InterfaceCRC: {1}", Value:=pDO^.SrcAdr, Value2:=InterfaceCRC);
                  end_if;
                end_if;
                // path can exist only once in a system
                return;
              elsif (pHelpPdo^.PdoInfo.Info.VirtualPDOsCreated = FALSE) then
                // it's a broadcast, the IF-CRC matches and we didn't create virtual PDOs so far
                pHelpSafety := pFirstSafetyComponent;
                while pHelpSafety do
                  if (pHelpPdo^.PdoInfo.pSourcePath^ = pHelpSafety^.pPath^) &
                     (To_StdLib.MemCmp(pHelpSafety^.pPath + 1, pHelpPdo^.PdoInfo.pSourcePath + 2 + pHelpPdo^.PdoInfo.pSourcePath^ - pHelpSafety^.pPath^, pHelpSafety^.pPath^) = 0) then

                    // change the command, because now we forward it to the receiver
                    pPara^.uiCmd := CMD_SM_SDO_TO_MODULE;

                    pHelpSafety^.pThis^.NewInst(pPara, #MyResult);
                    return;
                  else
                    pHelpSafety := pHelpSafety^.pNext;
                  end_if;
                end_while;
              end_if;
            end_if;

            pHelpPdo := pHelpPdo^.pNext;
          end_while;

          pHelpConfig := pHelpConfig^.pNext;
        end_while;
      end_if;
    end_if;

    // check if there is any interface frame domain optional and not available
    pHelpManaging := pFirstManagingInterfaceComponent;
    while pHelpManaging do
      if (pHelpManaging^.InfoBits.IsSynchron = 0) & (pHelpManaging^.InfoBits.IsOptional = 1) then
        // found one => no error here
        return;
      end_if;

      pHelpManaging := pHelpManaging^.pNext;
    end_while;

    // no optional interface domains missing => must be an error
    LogError("@0468 (SafetyManager::CheckTopSDO) Couldn't find InterfaceCRC. Check SafetyDesigner projects, maybe the interface variables do not match.");
    LogValue("SrcAddr: {0} / InterfaceCRC: {1}", Value:=pDO^.SrcAdr, Value2:=InterfaceCRC);
    ClassState := -8;

  // check if it's a local interface frame and we have no interface frame domains
  elsif (pCompDestPath^ = INTERFACE_CRC_MODE) then
    // after the mode byte we find the interface CRC
    InterfaceCRC := ((pCompDestPath + 1)$^HDINT)^;

    // search for the CRC
    pHelpSafety := NIL;
    if LocalIFNo then
      for i := 0 to (LocalIFNo-1) do
        if aLocalIFs[i].InterfaceCRC = InterfaceCRC then
          // found it
          pHelpSafety := aLocalIFs[i].pSafetyModule;
          exit;
        end_if;
      end_for;
    end_if;

    if pHelpSafety then
      // change the command, because now we forward it to the receiver
      pPara^.uiCmd := CMD_SM_SDO_TO_MODULE;

      pHelpSafety^.pThis^.NewInst(pPara, #MyResult);
    else
      // check the slave modules if there is one with the interface frame we need
      TargetSafetyNbr := 0;
      pHelpConfig := pConfigs;
      while pHelpConfig do
        pHelpSlave := pHelpConfig^.pFirstSlaveCfg;
        while pHelpSlave do

          if (pHelpSlave^.SlaveInfo.Info.IsInterface) & (pHelpSlave^.SlaveInfo.InterfaceCRC = InterfaceCRC) then
            // we have to add some additional information to the message

            (*
              Memory structure:
                1 Byte destination domain
                1 Byte IsInterfaceFrame (0/1)
                2 Byte length of uncompressed path
                x Byte uncompressed path
                x Byte SDO message
            *)

            MyPara.uiCmd := CMD_SM_TOP_SDO_TO_MODULE;
            MyPara.aPara[0] := sizeof(USINT) + sizeof(BOOL) + sizeof(UINT) + pHelpSlave^.SlaveInfo.PathLen + pPara^.aPara[0];

            if ud_SizeTempMemCy >= MyPara.aPara[0]$UDINT then
              pTempMem := pTempMemCy$^USINT;
            else
              LogError("@0440 (SafetyManager::CheckTopSDO) Temporary memory for cyclic task is too small!");
              LogValue("AvaliableMem: {0} / NeededMem: {1}", Value:=ud_SizeTempMemCy, Value2:=MyPara.aPara[0]$UDINT);
              return;
            end_if;

            TmpLen := pHelpSlave^.SlaveInfo.PathLen; // save some time with this local variable
            DomainChangeFound := FALSE;
            pHelp := pHelpSlave^.SlaveInfo.pPath + TmpLen - 2; // pointer on penultimate byte of path
            // search from the end for the last domain change
            for i := (TmpLen-2) to 3 by -1 do
              if pHelp^ = HWT_ESCAPE_DOMAIN then
                DomainChangeFound := TRUE;
                DestDomain := (pHelp + 1)^;
                exit;
              end_if;

              pHelp -= sizeof(USINT);
            end_for;

            // if there was no domainchange
            if DomainChangeFound = FALSE then
              // the master is the Dest
              DestDomain := (pHelpSlave^.SlaveInfo.pPath + 2)^;
            end_if;

            pHelp := pTempMem;

            // destination domain
            pHelp^ := DestDomain;
            pHelp += sizeof(USINT);

            // is it for an interface frame?
            pHelp^$BOOL := TRUE;
            pHelp += sizeof(BOOL);

            // length of uncompressed path
            pHelp^$UINT := TmpLen;
            pHelp += sizeof(UINT);

            // uncompressed path
            _memcpy(ptr1:=pHelp, ptr2:=pHelpSlave^.SlaveInfo.pPath, cntr:=TmpLen);
            pHelp += TmpLen;

            // SDO message
            _memcpy(ptr1:=pHelp, ptr2:=pDO, cntr:=pPara^.aPara[0]$UDINT);

            MyPara.aPara[1] := pTempMem$DINT;

            NewInst(#MyPara, #MyResult);

            // path can exist only once in a system
            return;
          end_if;

          pHelpSlave := pHelpSlave^.pNext;
        end_while;

        pHelpModule := pHelpConfig^.pFirstModuleCfg;
        while pHelpModule do
          if pHelpModule^.ModuleInfo.InterfaceCRC = InterfaceCRC then
            // if we found our target => forward the SDO to it
            TargetSafetyNbr := pHelpModule^.ModuleInfo.SafetyNbr;

            pHelpSafety := pFirstSafetyComponent;
            while pHelpSafety do
              // we compare the safety number
              if pHelpSafety^.SafetyNbr = TargetSafetyNbr then
                // change the command, because now we forward it to the receiver
                pPara^.uiCmd := CMD_SM_SDO_TO_MODULE;

                pHelpSafety^.pThis^.NewInst(pPara, #MyResult);

                return;
              end_if;

              pHelpSafety := pHelpSafety^.pNext;
            end_while;
          end_if;

          pHelpModule := pHelpModule^.pNext;
        end_while;

        pHelpConfig := pHelpConfig^.pNext;
      end_while;

      LogError("@046D (SafetyManager::CheckTopSDO) Couldn't find target of SDO via TOP (Local Interface Frame)");
      LogValue("SrcAddr: {0} / InterfaceCRC: {1}", Value:=pDO^.SrcAdr, Value2:=InterfaceCRC);
    end_if;
  elsif (pCompDestPath^ = INTERFACE_IP_MODE) then

    IPAddr := ((pCompDestPath + 5)$^HDINT)^;
    // after the mode byte we find the interface CRC
    InterfaceCRC := ((pCompDestPath + 1)$^HDINT)^;

    // Check Valid IP address
    if IPAddr AND 16#00FFFFFF then

      if sUdpVars.ProducerConnectionNo then

      // check udp producer list (if available)
        pActConnection := #sUdpVars.paConnectionsToProducers^[0];
        for i := 0 to (sUdpVars.ProducerConnectionNo-1) do

          if pActConnection^.IFCRC = InterfaceCRC then
            // got it => forward the SDO
            TmpLen := pPara^.aPara[0]$UINT;

            if TmpLen <= UDP_MAX_SDO_SIZE then
              // check for unsent SDO first
              if pActConnection^.ActSendData.SdoLength = 0 then
                UdpSendData.SectionStart();

                _memcpy(ptr1:=#pActConnection^.ActSendData.SdoData, ptr2:=pPara^.aPara[1]$pVoid, cntr:=TmpLen);
                pActConnection^.ActSendData.SdoLength     := TmpLen$USINT;

                UdpSendData.SectionStop();
              else
                sUdpVars.SdoAlreadyUsedCnt += 1;
              end_if;
            else
              LogError("@046E (SafetyManager::CheckTopSDO) SDO size exceeds the allowed size (Compressed Topology Path: UDP)");
            end_if;

            return;
          end_if;

          pActConnection += sizeof(t_UdpConnection);
        end_for;
      end_if;

      LogError("@146F (SafetyManager::CheckTopSDO) Couldn't find destination of SDO. (Compressed Topology Path: UDP)");
      LogValue("SrcAddr: {0} / InterfaceCRC: {1}", Value:=pDO^.SrcAdr, Value2:=((pCompDestPath + 1)$^HDINT)^);
    else

      // if source is in this station => search for managing components to forward
      pHelpSafety := pFirstSafetyComponent;

      while pHelpSafety do

        if pHelpSafety^.SafetyNbr = pDO^.SrcAdr then
          exit;
        end_if;

        pHelpSafety := pHelpSafety^.pNext;
      end_while;

      if pHelpSafety then

        // We are soure, send the data
        pHelpManaging := pFirstManagingInterfaceComponent;

        while pHelpManaging do

          if pHelpManaging^.pModulePath & pHelpManaging^.pModulePath^ = 3 then

            if ( (pHelpManaging^.pModulePath + 3)^ = HWT_ESCAPE_SAFETY_CUSTOM) &
                 (pHelpManaging^.pModulePath + 4)^ = (IPAddr shr 24)$USINT   then

              if pHelpManaging^.InfoBits.IsSynchron then
                pHelpManaging^.pThis^.NewInst(pPara, #MyResult);
              end_if;

              return;
            end_if;

          end_if;

          pHelpManaging := pHelpManaging^.pNext;
        end_while;

      else // source not here => search for destination with IF CRC

        // check if we have a module with this path
        pHelpConfig := pConfigs;
        while pHelpConfig do

          pHelpModule := pHelpConfig^.pFirstModuleCfg;
          while pHelpModule do
            if pHelpModule^.ModuleInfo.InterfaceCRC = InterfaceCRC then
              // if we found our target => forward the SDO to it
              TargetSafetyNbr := pHelpModule^.ModuleInfo.SafetyNbr;

              pHelpSafety := pFirstSafetyComponent;
              while pHelpSafety do
                // we compare the safety number
                if pHelpSafety^.SafetyNbr = TargetSafetyNbr then
                  // change the command, because now we forward it to the receiver
                  pPara^.uiCmd := CMD_SM_SDO_TO_MODULE;

                  pHelpSafety^.pThis^.NewInst(pPara, #MyResult);

                  return;
                end_if;

                pHelpSafety := pHelpSafety^.pNext;
              end_while;
            end_if;

            pHelpModule := pHelpModule^.pNext;
          end_while;

          pHelpConfig := pHelpConfig^.pNext;
        end_while;

      end_if;

      LogValue("@0471 (SafetyManager::CheckTopSDO) Couldn't find destination of SDO. (Custom connection no: {0})", Value:=(IPAddr shr 24) );
      LogValue("SrcAddr: {0} / InterfaceCRC: {1}", Value:=pDO^.SrcAdr, Value2:=((pCompDestPath + 1)$^HDINT)^);

    end_if;
  else
    // check if we have a module with this path
    pHelpConfig := pConfigs;
    while pHelpConfig do
      pHelpModule := pHelpConfig^.pFirstModuleCfg;
      while pHelpModule do
        if (To_StdLib.MemCmp(pCompDestPath, pHelpModule^.ModuleInfo.pCompPath, pHelpModule^.ModuleInfo.CompPathLen) = 0) then
          // we have to add some additional information to the message

          (*
            Memory structure:
              1 Byte destination domain
              1 Byte IsInterfaceFrame (0/1)
              2 Byte length of uncompressed path
              x Byte uncompressed path
              x Byte SDO message
          *)

          TmpLen := pHelpModule^.ModuleInfo.PathLen; // save some time with this local variable
          MyPara.uiCmd := CMD_SM_TOP_SDO_TO_MODULE;
          MyPara.aPara[0] := sizeof(USINT) + sizeof(BOOL) + sizeof(UINT) + TmpLen + pPara^.aPara[0];
          if ud_SizeTempMemCy >= MyPara.aPara[0]$UDINT then
            pTempMem := pTempMemCy$^USINT;
          else
            LogError("@0440 (SafetyManager::CheckTopSDO) Temporary memory for cyclic task is too small!");
            LogValue("AvaliableMem: {0} / NeededMem: {1}", Value:=ud_SizeTempMemCy, Value2:=MyPara.aPara[0]$UDINT);
            return;
          end_if;

          DomainChangeFound := FALSE;
          pHelp := pHelpModule^.ModuleInfo.pPath + TmpLen - 2; // pointer on penultimate byte of path
          // search from the end for the last domain change
          for i := (TmpLen-2) to 3 by -1 do
            if pHelp^ = HWT_ESCAPE_DOMAIN then
              DomainChangeFound := TRUE;
              DestDomain := (pHelp + 1)^;
              exit;
            end_if;

            pHelp -= sizeof(USINT);
          end_for;

          // if there was no domainchange
          if DomainChangeFound = FALSE then
            // the master is the Dest
            DestDomain := (pHelpModule^.ModuleInfo.pPath + 2)^;
          end_if;

          pHelp := pTempMem;

          // destination domain
          pHelp^ := DestDomain;
          pHelp += sizeof(USINT);

          // is it for an interface frame?
          pHelp^$BOOL := FALSE;
          pHelp += sizeof(BOOL);

          // length of uncompressed path
          pHelp^$UINT := TmpLen;
          pHelp += sizeof(UINT);

          // uncompressed path
          _memcpy(ptr1:=pHelp, ptr2:=pHelpModule^.ModuleInfo.pPath, cntr:=TmpLen);
          pHelp += TmpLen;

          // SDO message
          _memcpy(ptr1:=pHelp, ptr2:=pDO, cntr:=pPara^.aPara[0]$UDINT);

          MyPara.aPara[1] := pTempMem$DINT;

          NewInst(#MyPara, #MyResult);

          // path can exist only once in a system
          return;
        end_if;

        pHelpModule := pHelpModule^.pNext;
      end_while;

      if pHelpConfig^.SafetyNbr = pDO^.SrcAdr then
        pHelpSlave := pHelpConfig^.pFirstSlaveCfg;
        while pHelpSlave do
          if (To_StdLib.MemCmp(pCompDestPath, pHelpSlave^.SlaveInfo.pCompPath, pHelpSlave^.SlaveInfo.CompPathLen) = 0) then
            // we have to add some additional information to the message

            (*
              Memory structure:
                1 Byte destination domain
                1 Byte IsInterfaceFrame (0/1)
                2 Byte length of uncompressed path
                x Byte uncompressed path
                x Byte SDO message
            *)

            TmpLen := pHelpSlave^.SlaveInfo.PathLen; // save some time with this local variable
            MyPara.uiCmd := CMD_SM_TOP_SDO_TO_MODULE;
            MyPara.aPara[0] := sizeof(USINT) + sizeof(BOOL) + sizeof(UINT) + TmpLen + pPara^.aPara[0];
            if ud_SizeTempMemCy >= MyPara.aPara[0]$UDINT then
              pTempMem := pTempMemCy$^USINT;
            else
              LogError("@0440 (SafetyManager::CheckTopSDO) Temporary memory for cyclic task is too small!");
              LogValue("AvaliableMem: {0} / NeededMem: {1}", Value:=ud_SizeTempMemCy, Value2:=MyPara.aPara[0]$UDINT);
              return;
            end_if;

            DomainChangeFound := FALSE;
            pHelp := pHelpSlave^.SlaveInfo.pPath + TmpLen - 2; // pointer on penultimate byte of path
            // search from the end for the last domain change
            for i := (TmpLen-2) to 3 by -1 do
              if pHelp^ = HWT_ESCAPE_DOMAIN then
                DomainChangeFound := TRUE;
                DestDomain := (pHelp + 1)^;
                exit;
              end_if;

              pHelp -= sizeof(USINT);
            end_for;

            // if there was no domainchange
            if DomainChangeFound = FALSE then
              // the master is the Dest
              DestDomain := (pHelpSlave^.SlaveInfo.pPath + 2)^;
            end_if;

            pHelp := pTempMem;

            // destination domain
            pHelp^ := DestDomain;
            pHelp += sizeof(USINT);

            // is it for an interface frame?
            pHelp^$BOOL := FALSE;
            pHelp += sizeof(BOOL);

            // length of uncompressed path
            pHelp^$UINT := TmpLen;
            pHelp += sizeof(UINT);

            // uncompressed path
            _memcpy(ptr1:=pHelp, ptr2:=pHelpSlave^.SlaveInfo.pPath, cntr:=TmpLen);
            pHelp += TmpLen;

            // SDO message
            _memcpy(ptr1:=pHelp, ptr2:=pDO, cntr:=pPara^.aPara[0]$UDINT);

            MyPara.aPara[1] := pTempMem$DINT;

            NewInst(#MyPara, #MyResult);

            // path can exist only once in a system
            return;
          end_if;

          pHelpSlave := pHelpSlave^.pNext;
        end_while;
      end_if;

      pHelpConfig := pHelpConfig^.pNext;
    end_while;

    LogError("@0472 (SafetyManager::CheckTopSDO) Couldn't find destination of SDO. (Compressed Topology Path)");
    LogValue("SrcAddr: {0} / InterfaceCRC: {1}", Value:=pDO^.SrcAdr, Value2:=((pCompDestPath + 1)$^HDINT)^);

  end_if;

END_FUNCTION

FUNCTION SafetyManager::TopSDODest
  VAR_INPUT
    pPara 	: ^CmdStruct;
    pResult 	: ^results;
  END_VAR
  VAR_OUTPUT
    IsDestDomain 	: BOOL;
  END_VAR
  VAR
    pHelpUSINT : ^USINT;
    PathLength : UINT;
    pPath : ^USINT;
    pHelpSafety : ^t_SafetyComponent;
  END_VAR

  IsDestDomain := FALSE;
(*
  Memory structure:
    1 Byte destination domain
    1 Byte IsInterfaceFrame (0/1)
    2 Byte length of uncompressed path
    x Byte uncompressed path
    x Byte SDO message
*)

  // check size (at least 1 byte for the destination domain + 2 byte for the path length + the header of the SDO message)
  if pPara^.aPara[0] > (sizeof(USINT) + sizeof(PathLength) + sizeof(SafetyCDIAS_Base::SDOHeader.StdHeader)) then
    pHelpUSINT := (pPara^.aPara[1])$^USINT;

    // domain
    pHelpUSINT += sizeof(USINT);

    // is it an interface frame info?
    pHelpUSINT += sizeof(BOOL);

    // path length
    PathLength := (pHelpUSINT$^UINT)^;
    pHelpUSINT += sizeof(UINT);

    // path
    pPath := pHelpUSINT;
    pHelpUSINT += PathLength;

    // pHelpUSINT points now to the SDO message

    // now we search the logged in modules for one with a matching topology path
    if pFirstSafetyComponent then

      pHelpSafety := pFirstSafetyComponent;
      while pHelpSafety do
        // we compare the last x byte (where x is the length of the local path including the domain) => update: no more transfer between different domains,
        //                                                                                                      therefore the length has to match before we compare the end of the path
        if pHelpSafety^.pPath & (pHelpSafety^.pPath^ = pPath^) & (To_StdLib.MemCmp(pHelpSafety^.pPath + 1, pPath + 2 + pPath^ - pHelpSafety^.pPath^, pHelpSafety^.pPath^) = 0) then
          pPara^.uiCmd := CMD_SM_SDO_TO_MODULE;
          pPara^.aPara[0] := pPara^.aPara[0] - (sizeof(USINT) + sizeof(PathLength) + PathLength);
          pPara^.aPara[1] := pHelpUSINT$DINT;

          pHelpSafety^.pThis^.NewInst(pPara, pResult);

          IsDestDomain := TRUE;
          return;
        end_if;

        pHelpSafety := pHelpSafety^.pNext;
      end_while;
    end_if;
  end_if;

END_FUNCTION

FUNCTION SafetyManager::PDOLengthCorrection
  VAR
    pHelpConfig : ^t_CfgListElem;
    pHelpPDO    : ^t_PdoListElem;
    pHelpModule : ^t_ModuleListElem;
    pHelpSearchConfig : ^t_CfgListElem;
    FoundIt : BOOL;
    GotFirst : BOOL;
  END_VAR

  // with FSoE we use connections instead of the PDOs (PDOs are only remembered to check the optional state)
  if b_GotFSoEModules then
    return;
  end_if;

  GotFirst := FALSE;

  // check if there is a PDO with a zero length
  pHelpConfig := pConfigs;
  while pHelpConfig do
    pHelpPDO := pHelpConfig^.pFirstPdoCfg;
    while pHelpPDO do
      // remember the first PDO found as our act (to start from)
      if GotFirst = FALSE then
        GotFirst := TRUE;

        pActualSendCfg := pHelpConfig;
        pActualSendPDO := pHelpPDO;
      end_if;

      // if there is a PDO with no length
      if pHelpPDO^.PdoInfo.PdoLen = 0 then
        FoundIt := FALSE;
        pHelpSearchConfig := pConfigs;
        // search for the source module, because we use the length of it
        while pHelpSearchConfig & (FoundIt = FALSE) do
          pHelpModule := pHelpSearchConfig^.pFirstModuleCfg;
          while pHelpModule & (FoundIt = FALSE) do
            if pHelpModule^.ModuleInfo.PathLen = pHelpPDO^.PdoInfo.SourcePathLen then
              if (To_StdLib.MemCmp(pHelpModule^.ModuleInfo.pPath, pHelpPDO^.PdoInfo.pSourcePath, pHelpModule^.ModuleInfo.PathLen) = 0) then
                pHelpPDO^.PdoInfo.PdoLen := pHelpModule^.ModuleInfo.PdoOutLen;
                FoundIt := TRUE;
              end_if;
            end_if;

            pHelpModule := pHelpModule^.pNext;
          end_while;

          pHelpSearchConfig := pHelpSearchConfig^.pNext;
        end_while;
      end_if;

      pHelpPDO := pHelpPDO^.pNext;
    end_while;

    pHelpConfig := pHelpConfig^.pNext;
  end_while;

END_FUNCTION

FUNCTION SafetyManager::DoublePDOEntry
  VAR_INPUT
    NewPDO 	: t_PdoCfg;
    pNewCfg 	: ^t_CfgListElem;
  END_VAR
  VAR_OUTPUT
    IsDoubleEntry 	: BOOL;
  END_VAR
  VAR
    pHelpCfg : ^t_CfgListElem;
    pHelpPdo : ^t_PdoListElem;
  END_VAR

  IsDoubleEntry := FALSE;

  // if it's our first config, there is no chance for a double PDO => check only if not first config
  if pNewCfg <> pConfigs then
    // otherwise: search all prior configs for the same PDO (source and destination path match)
    pHelpCfg := pConfigs;
    while pHelpCfg <> pNewCfg do
      pHelpPdo := pHelpCfg^.pFirstPdoCfg;
      while pHelpPdo do
        if (pHelpPdo^.PdoInfo.SourcePathLen = NewPDO.SourcePathLen) & (pHelpPdo^.PdoInfo.DestPathLen = NewPDO.DestPathLen) &
           (To_StdLib.MemCmp(pHelpPdo^.PdoInfo.pSourcePath, NewPDO.pSourcePath, NewPDO.SourcePathLen) = 0) &
           (To_StdLib.MemCmp(pHelpPdo^.PdoInfo.pDestPath, NewPDO.pDestPath, NewPDO.DestPathLen) = 0) then
          // we found the same PDO in a prior config
          IsDoubleEntry := TRUE;
          return;
        end_if;

        pHelpPdo := pHelpPdo^.pNext;
      end_while;

      pHelpCfg := pHelpCfg^.pNext;
    end_while;
  end_if;

END_FUNCTION

FUNCTION SafetyManager::StoreInterfaceRoutingList
  VAR_INPUT
    pPara 	: ^CmdStruct;
    pResult 	: ^results;
    IsFSoE 	: BOOL;
  END_VAR
  VAR
    pHelpManaging : ^t_ManagingComponent;
    EntryNo       : USINT;
    i             : UDINT;
    pHelp         : ^t_InterfaceFrameInfo;
    ActOffset     : UDINT;
    pHelpFSoE     : ^t_IFConnectionInfo;
    j             : UDINT;
    GenerateNo    : USINT;
    OldFSoENo     : DINT;
  END_VAR

  if IsFSoE then

    // if we already have different data from this management component => delete the old stuff first
    if IFFSoENo then
      OldFSoENo := IFFSoENo$DINT;

      // remove the existing stuff of this managing component
      for i$DINT := (OldFSoENo-1) to 0 by -1 do
        // check if it's from the same managing component
        if aIFFSoEInfos[i].pManaging^.pThis$DINT = pPara^.aPara[2] then
          // remove it

          // move the following blocks over this one (if it's not the last)
          if i$UDINT < IFFSoENo-1 then
            for j := i to (IFFSoENo-2) do
              aIFFSoEInfos[j] := aIFFSoEInfos[j+1];
            end_for;
          end_if;
          IFFSoENo -= 1;
        end_if;
      end_for;
    end_if;

    EntryNo := ((pPara^.aPara[0] - sizeof(t_IFInfoFSoE.IsResponse)) / sizeof(t_IFConnectionInfo))$USINT;
    if (EntryNo + IFFSoENo <= MAX_MODULES_IN_OTHER_DOMAINS) then
      ActOffset := 0;
      pHelpManaging := pFirstManagingInterfaceComponent;
      while pHelpManaging do
        // if we found the sender of this list in our list of interfaceframe components, remember the safety numbers
        if pHelpManaging^.pThis$DINT = pPara^.aPara[2] then
          if EntryNo then

            // set the help pointer to the first entry of the interface frame info array
            pHelpFSoE := pPara^.aPara[1]$^t_IFConnectionInfo + sizeof(BOOL);
            for i := 0 to (EntryNo-1) do
              pHelpManaging^.ModuleInfo[i].SafetyNbr := pHelpFSoE^.SafetyNbr;

              if pHelpFSoE^.Flags.IsMaster then
                pHelpManaging^.ModuleInfo[i].InfoBits.IsFSoEMaster := TRUE;
                pHelpManaging^.ModuleInfo[i].InfoBits.IsFSoESlave  := FALSE;
              else
                pHelpManaging^.ModuleInfo[i].InfoBits.IsFSoEMaster := FALSE;
                pHelpManaging^.ModuleInfo[i].InfoBits.IsFSoESlave  := TRUE;
              end_if;

              // we save the whole info for PDO/SDO routing
              aIFFSoEInfos[IFFSoENo].FromOtherSide := pHelpFSoE^;
              aIFFSoEInfos[IFFSoENo].FromOtherSide.FollowUps := 0; // only relevant for the transfer to this domain
              aIFFSoEInfos[IFFSoENo].pManaging := pHelpManaging;

              IFFSoENo += 1;

              if pHelpFSoE^.FollowUps then
                GenerateNo := pHelpFSoE^.FollowUps;
                for j := 1 to GenerateNo do
                  // we save the whole info for PDO/SDO routing
                  aIFFSoEInfos[IFFSoENo].FromOtherSide := pHelpFSoE^;
                  aIFFSoEInfos[IFFSoENo].FromOtherSide.FollowUps := 0; // only relevant for the transfer to this domain
                  aIFFSoEInfos[IFFSoENo].pManaging := pHelpManaging;

                  IFFSoENo += 1;
                end_for;
              end_if;

              pHelpFSoE += sizeof(t_IFConnectionInfo);
            end_for;
          end_if;

          pHelpManaging^.ModuleNo := EntryNo;

          pHelpManaging^.InfoBits.GotIFInfo := TRUE;
          return;
        end_if;

        pHelpManaging := pHelpManaging^.pNext;
      end_while;
    else
      LogError("@0473 (SafetyManager::StoreInterfaceRoutingList) Invalid size of configuration (FSoE)");
    end_if;
  else
    EntryNo := ((pPara^.aPara[0] - sizeof(t_IFInfo.IsResponse)) / sizeof(t_InterfaceFrameInfo))$USINT;

    if (EntryNo + InterfaceFrameNo <= MAX_MODULES_IN_OTHER_DOMAINS) then
      ActOffset := 0;
      pHelpManaging := pFirstManagingInterfaceComponent;
      while pHelpManaging do
        // if we found the sender of this list in our list of interfaceframe components, remember the safety numbers
        if pHelpManaging^.pThis$DINT = pPara^.aPara[2] then
          if EntryNo then
            // set the help pointer to the first entry of the interface frame info array
            pHelp := pPara^.aPara[1]$^t_InterfaceFrameInfo + sizeof(BOOL);
            for i := 0 to (EntryNo-1) do
              // we save the module info's with the domain interface module for TDO/SDO routing
              pHelpManaging^.ModuleInfo[i] := pHelp^.ModuleInfo;

              // we also save the whole info for PDO routing
              aInterfaceFrameInfos[InterfaceFrameNo] := pHelp^;

              // only for IFs where the communication partner is the source
              if aInterfaceFrameInfos[InterfaceFrameNo].IFPdoLen then
                aInterfaceFrameInfos[InterfaceFrameNo].OffsetInDomainModule := ActOffset;
                ActOffset += aInterfaceFrameInfos[InterfaceFrameNo].IFPdoLen;
              end_if;

              InterfaceFrameNo += 1;

              pHelp += sizeof(t_InterfaceFrameInfo);
            end_for;
          end_if;

          pHelpManaging^.ModuleNo := EntryNo;

          pHelpManaging^.InfoBits.GotIFInfo := TRUE;
          return;
        end_if;

        pHelpManaging := pHelpManaging^.pNext;
      end_while;
    else
      LogError("@0475 (SafetyManager::StoreInterfaceRoutingList) Invalid size of configuration");
    end_if;
  end_if;

END_FUNCTION

FUNCTION SafetyManager::AllInterfaceCfgsArrived
  VAR_OUTPUT
    AllReady 	: BOOL;
  END_VAR
  VAR
    pHelpManaging : ^t_ManagingComponent;
  END_VAR

  AllReady := TRUE;

  // check if we have the safety numbers for every interface managing module in the system
  pHelpManaging := pFirstManagingInterfaceComponent;
  while pHelpManaging do
    if pHelpManaging^.InfoBits.IsSynchron & (pHelpManaging^.InfoBits.GotIFInfo = FALSE) then
      AllReady := FALSE;
      return;
    end_if;

    pHelpManaging := pHelpManaging^.pNext;
  end_while;

END_FUNCTION

FUNCTION SafetyManager::SendInterfaceConfigs
  VAR_INPUT
    DestinationThis 	: pVirtualBase;(* := NIL *)
    IsResponse 	: BOOL;(* := FALSE *)
    IsFSoE 	: BOOL;
  END_VAR
  VAR
    pHelpCfg                  : ^t_CfgListElem;
    pHelpModule               : ^t_ModuleListElem;
    pHelpPdo                  : ^t_PdoListElem;
    pHelpConnection           : ^t_FSoEConnectionDetails;
    MyPara                    : CmdStruct;
    MyResult                  : results;
    TmpIFInfo                 : t_IFInfo;
    ModuleInfoNo              : USINT;
    i                         : UDINT;
    pActCRC                   : ^HDINT;
    TmpIFConn                 : t_IFInfoFSoESend;
    pLastReferenceConnection  : ^t_IFConnectionInfo;
  END_VAR

  // collect the safety numbers of this system
  ModuleInfoNo := 0;

  if IsFSoE then
    //reset memory => now 0 is an invalid safety number (= unused element of the array)
    _memset(dest:=#TmpIFConn, usByte:=0, cntr:=sizeof(t_IFInfoFSoESend));
    TmpIFConn.IsResponse := IsResponse;

    pLastReferenceConnection  := NIL;

    // if not all configs available, create and send the available data
    if (LocalCPUCfgNo <> LocalCPUNo) then
      // check FSoE Connections in the available configs
      pHelpCfg := pConfigs;
      while pHelpCfg do
        pHelpConnection := pHelpCfg^.pFirstFSoEConnection;
        while pHelpConnection do
          // only interface connections are relevant
          if pHelpConnection^.Flags.IsInterfaceConnection then
            if pLastReferenceConnection & (pHelpConnection^.SlaveAddress = pLastReferenceConnection^.SlaveAddress) &
               (pHelpConnection^.Flags.IsMaster = pLastReferenceConnection^.Flags.IsMaster) then
              pLastReferenceConnection^.FollowUps += 1;
            else
              // add the modules to the info message
              TmpIFConn.aConnectionInfos[ModuleInfoNo].Flags            := pHelpConnection^.Flags;
              TmpIFConn.aConnectionInfos[ModuleInfoNo].SlaveAddress     := pHelpConnection^.SlaveAddress;
              TmpIFConn.aConnectionInfos[ModuleInfoNo].SafetyNbr        := pHelpConnection^.OwnerSafetyNbr;
              TmpIFConn.aConnectionInfos[ModuleInfoNo].MasterReadSize   := pHelpConnection^.MasterReadSize;
              TmpIFConn.aConnectionInfos[ModuleInfoNo].MasterWriteSize  := pHelpConnection^.MasterWriteSize;
              TmpIFConn.aConnectionInfos[ModuleInfoNo].FollowUps        := 0;

              // some data are only available at the master
              if pHelpConnection^.Flags.IsMaster then
                // no follow ups for master connections
                pLastReferenceConnection                                := NIL;

                TmpIFConn.aConnectionInfos[ModuleInfoNo].ConnectionID   := pHelpConnection^.ConnectionID;
              else
                // update this value for the next connections with the same settings to save a lot of memory
                pLastReferenceConnection                                := #TmpIFConn.aConnectionInfos[ModuleInfoNo];

                TmpIFConn.aConnectionInfos[ModuleInfoNo].ConnectionID   := 0;
              end_if;

              if pHelpConnection^.SlavePathCompLen & pHelpConnection^.pSlavePathComp then
                TmpIFConn.aConnectionInfos[ModuleInfoNo].InterfaceCRC := (pHelpConnection^.pSlavePathComp$^HDINT + 1)^;
              else
                TmpIFConn.aConnectionInfos[ModuleInfoNo].InterfaceCRC := 0;
              end_if;

              ModuleInfoNo += 1;
            end_if;
          end_if;

          pHelpConnection := pHelpConnection^.pNext;
        end_while;

        pHelpCfg := pHelpCfg^.pNext;
      end_while;
    else
      // check FSoE Connections in the sorted list
      pHelpConnection := pSortedConnections;
      while pHelpConnection do
        // only interface connections are relevant
        if pHelpConnection^.Flags.IsInterfaceConnection then
          if pLastReferenceConnection & (pHelpConnection^.SlaveAddress = pLastReferenceConnection^.SlaveAddress) &
             (pHelpConnection^.Flags.IsMaster = pLastReferenceConnection^.Flags.IsMaster) then
            pLastReferenceConnection^.FollowUps += 1;
          else
            // add the modules to the info message
            TmpIFConn.aConnectionInfos[ModuleInfoNo].Flags            := pHelpConnection^.Flags;
            TmpIFConn.aConnectionInfos[ModuleInfoNo].SlaveAddress     := pHelpConnection^.SlaveAddress;
            TmpIFConn.aConnectionInfos[ModuleInfoNo].SafetyNbr        := pHelpConnection^.OwnerSafetyNbr;
            TmpIFConn.aConnectionInfos[ModuleInfoNo].MasterReadSize   := pHelpConnection^.MasterReadSize;
            TmpIFConn.aConnectionInfos[ModuleInfoNo].MasterWriteSize  := pHelpConnection^.MasterWriteSize;
            TmpIFConn.aConnectionInfos[ModuleInfoNo].FollowUps        := 0;

            // some data are only available at the master
            if pHelpConnection^.Flags.IsMaster then
              // no follow ups for master connections
              pLastReferenceConnection                                := NIL;

              TmpIFConn.aConnectionInfos[ModuleInfoNo].ConnectionID   := pHelpConnection^.ConnectionID;
            else
              // update this value for the next connections with the same settings to save a lot of memory
              pLastReferenceConnection                                := #TmpIFConn.aConnectionInfos[ModuleInfoNo];

              TmpIFConn.aConnectionInfos[ModuleInfoNo].ConnectionID   := 0;
            end_if;

            if pHelpConnection^.SlavePathCompLen & pHelpConnection^.pSlavePathComp then
              TmpIFConn.aConnectionInfos[ModuleInfoNo].InterfaceCRC := (pHelpConnection^.pSlavePathComp$^HDINT + 1)^;
            else
              TmpIFConn.aConnectionInfos[ModuleInfoNo].InterfaceCRC := 0;
            end_if;

            ModuleInfoNo += 1;
          end_if;
        end_if;

        pHelpConnection := pHelpConnection^.pNextSorted;
      end_while;
    end_if;

    CheckLocalSlaveAddresses();

    if b_AllLocalSlaveAddressesValid then
      MyPara.uiCmd := CMD_SM_IF_MODULE_INFO_FSOE_OK;
    else
      MyPara.uiCmd := CMD_SM_IF_MODULE_INFO_FSOE;
    end_if;

    MyPara.aPara[0] := ModuleInfoNo * sizeof(t_IFConnectionInfo) + sizeof(t_IFInfoFSoE.IsResponse);
    MyPara.aPara[1] := (#TmpIFConn)$DINT;
  else
    // browse through the configs
    TmpIFInfo.IsResponse := IsResponse;

    pHelpCfg := pConfigs;
    while pHelpCfg do
      pHelpPdo := pHelpCfg^.pFirstPdoCfg;
      while pHelpPdo do
        // if it's a interface broadcast
        if pHelpPdo^.PdoInfo.Info.IFBroadCast then
          // search for the source module
          pHelpModule := pHelpCfg^.pFirstModuleCfg;
          while pHelpModule do
            // if it's an interface source and the interface CRC matches the one of our PDO => Bingo! But to be sure we check also the path length and the path itself
            if pHelpModule^.ModuleInfo.Info.IsInterfaceSource & (pHelpModule^.ModuleInfo.InterfaceCRC = pHelpPdo^.PdoInfo.InterfaceCRC) &
              (pHelpModule^.ModuleInfo.PathLen = pHelpPdo^.PdoInfo.SourcePathLen) &
              (To_StdLib.MemCmp(pHelpModule^.ModuleInfo.pPath, pHelpPdo^.PdoInfo.pSourcePath, pHelpPdo^.PdoInfo.SourcePathLen) = 0) then

              TmpIFInfo.aModuleInfos[ModuleInfoNo].InterfaceCRC          := pHelpModule^.ModuleInfo.InterfaceCRC;
              TmpIFInfo.aModuleInfos[ModuleInfoNo].IFPdoLen              := pHelpPdo^.PdoInfo.PdoLen;
              TmpIFInfo.aModuleInfos[ModuleInfoNo].OffsetInDomainModule  := 0; // the correct offset is calculated in the receiver
              TmpIFInfo.aModuleInfos[ModuleInfoNo].ModuleInfo.SafetyNbr  := pHelpModule^.ModuleInfo.SafetyNbr;
